Universal Robots URScript: FaiChun_9 Jan_7.script

def Machining1():
  # Default parameters:
  global speed_ms = 0.1
  global speed_rads = 0.75
  global accel_mss = 3
  global accel_radss = 1.2
  global blend_radius_m = 0.0002

  # Add subprograms here
  # Start of main program
  # Program generated by RoboDK v5.6.8 for UR10e on 10/01/2025 13:02:06
  # Using nominal kinematics.
  blend_radius_m = 0.0002
  speed_ms = 0.1
  # set_reference(p[0.355000, -0.055000, 0.001500, 0.000000, 0.000000, 0.000000])
  set_tcp(p[0.000000, 0.000000, 0.252000, 0.000000, 0.000000, 0.000000])
  # Show Tool
  movej([0.687885, -1.099321, -2.618738, -0.994329, 1.570796, 2.258681],accel_radss,speed_rads,0,blend_radius_m)
  movel([0.687885, -1.158787, -2.657718, -0.895884, 1.570796, 2.258681],accel_mss,speed_ms,0,blend_radius_m)
  #SetTool1
  #M_RunCode6
  #SetRPM60000
  speed_ms = 0.1
  #M_RunCode3
  movel([0.687885, -1.186172, -2.672546, -0.853671, 1.570796, 2.258681],accel_mss,speed_ms,0,blend_radius_m)
  speed_ms = 0.003
  movel([0.687885, -1.193386, -2.676190, -0.842813, 1.570796, 2.258681],accel_mss,speed_ms,0,blend_radius_m)
  speed_ms = 0.007
  movel([0.511185, -1.481281, -2.488242, -0.742866, 1.570796, 2.081982],accel_mss,speed_ms,0,blend_radius_m)
  movel([0.262250, -1.477063, -2.491849, -0.743477, 1.570796, 1.833046],accel_mss,speed_ms,0,blend_radius_m)
  movel([0.358500, -1.184451, -2.680352, -0.847585, 1.570796, 1.929297],accel_mss,speed_ms,0,blend_radius_m)
  movel([0.687885, -1.193386, -2.676190, -0.842813, 1.570796, 2.258681],accel_mss,speed_ms,0,blend_radius_m)
  speed_ms = 0.003
  movel([0.687885, -1.186172, -2.672546, -0.853671, 1.570796, 2.258681],accel_mss,speed_ms,0,blend_radius_m)
  speed_ms = 0.1
  movel([0.687885, -1.158787, -2.657718, -0.895884, 1.570796, 2.258681],accel_mss,speed_ms,0,blend_radius_m)
  #M_RunCode9
  movel([0.673659, -1.163346, -2.655655, -0.893388, 1.570796, 2.244455],accel_mss,speed_ms,0,blend_radius_m)
  #M_RunCode3
  movel([0.673659, -1.190701, -2.670423, -0.851265, 1.570796, 2.244455],accel_mss,speed_ms,0,blend_radius_m)
  speed_ms = 0.003
  movel([0.673659, -1.197905, -2.674052, -0.840433, 1.570796, 2.244455],accel_mss,speed_ms,0,blend_radius_m)
  speed_ms = 0.007
  movel([0.670159, -1.203367, -2.671437, -0.837585, 1.570796, 2.240955],accel_mss,speed_ms,0,blend_radius_m)
  movel([0.674542, -1.204354, -2.670961, -0.837074, 1.570796, 2.245338],accel_mss,speed_ms,0,blend_radius_m)
  movel([0.669404, -1.212334, -2.667074, -0.832981, 1.570796, 2.240200],accel_mss,speed_ms,0,blend_radius_m)
  movel([0.665043, -1.211367, -2.667549, -0.833473, 1.570796, 2.235840],accel_mss,speed_ms,0,blend_radius_m)
  movel([0.663268, -1.214147, -2.666181, -0.832061, 1.570796, 2.234065],accel_mss,speed_ms,0,blend_radius_m)
  movel([0.667621, -1.215107, -2.665706, -0.831575, 1.570796, 2.238418],accel_mss,speed_ms,0,blend_radius_m)
  movel([0.663402, -1.221682, -2.662429, -0.828278, 1.570796, 2.234198],accel_mss,speed_ms,0,blend_radius_m)
  movel([0.662590, -1.222948, -2.661792, -0.827649, 1.570796, 2.233387],accel_mss,speed_ms,0,blend_radius_m)
  movel([0.656171, -1.221563, -2.662488, -0.828337, 1.570796, 2.226968],accel_mss,speed_ms,0,blend_radius_m)
  movel([0.659538, -1.216260, -2.665135, -0.830994, 1.570796, 2.230334],accel_mss,speed_ms,0,blend_radius_m)
  movel([0.657269, -1.215780, -2.665373, -0.831236, 1.570796, 2.228065],accel_mss,speed_ms,0,blend_radius_m)
  movel([0.652180, -1.223829, -2.661348, -0.827212, 1.570796, 2.222977],accel_mss,speed_ms,0,blend_radius_m)
  movel([0.660845, -1.225674, -2.660415, -0.826300, 1.570796, 2.231641],accel_mss,speed_ms,0,blend_radius_m)
  movel([0.581204, -1.353206, -2.585789, -0.773394, 1.570796, 2.152000],accel_mss,speed_ms,0,blend_radius_m)
  movel([0.518903, -1.459211, -2.506807, -0.746371, 1.570796, 2.089699],accel_mss,speed_ms,0,blend_radius_m)
  movel([0.511689, -1.458211, -2.507631, -0.746547, 1.570796, 2.082486],accel_mss,speed_ms,0,blend_radius_m)
  movel([0.508628, -1.463700, -2.503092, -0.745597, 1.570796, 2.079424],accel_mss,speed_ms,0,blend_radius_m)
  movel([0.510492, -1.463952, -2.502883, -0.745554, 1.570796, 2.081288],accel_mss,speed_ms,0,blend_radius_m)
  movel([0.512509, -1.460346, -2.505871, -0.746172, 1.570796, 2.083305],accel_mss,speed_ms,0,blend_radius_m)
  movel([0.517829, -1.461092, -2.505254, -0.746043, 1.570796, 2.088625],accel_mss,speed_ms,0,blend_radius_m)
  movel([0.517338, -1.461959, -2.504537, -0.745893, 1.570796, 2.088135],accel_mss,speed_ms,0,blend_radius_m)
  movel([0.514822, -1.466415, -2.500830, -0.745144, 1.570796, 2.085618],accel_mss,speed_ms,0,blend_radius_m)
  movel([0.511249, -1.465915, -2.501248, -0.745226, 1.570796, 2.082045],accel_mss,speed_ms,0,blend_radius_m)
  movel([0.510209, -1.467774, -2.499694, -0.744921, 1.570796, 2.081005],accel_mss,speed_ms,0,blend_radius_m)
  movel([0.513778, -1.468272, -2.499276, -0.744840, 1.570796, 2.084574],accel_mss,speed_ms,0,blend_radius_m)
  movel([0.510816, -1.473540, -2.494840, -0.744009, 1.570796, 2.081613],accel_mss,speed_ms,0,blend_radius_m)
  movel([0.507266, -1.473049, -2.495255, -0.744085, 1.570796, 2.078063],accel_mss,speed_ms,0,blend_radius_m)
  movel([0.505298, -1.476588, -2.492253, -0.743548, 1.570796, 2.076095],accel_mss,speed_ms,0,blend_radius_m)
  movel([0.500042, -1.475891, -2.492846, -0.743652, 1.570796, 2.070838],accel_mss,speed_ms,0,blend_radius_m)
  movel([0.501993, -1.472345, -2.495850, -0.744194, 1.570796, 2.072789],accel_mss,speed_ms,0,blend_radius_m)
  movel([0.500139, -1.472105, -2.496053, -0.744231, 1.570796, 2.070935],accel_mss,speed_ms,0,blend_radius_m)
  movel([0.498194, -1.475653, -2.493048, -0.743688, 1.570796, 2.068990],accel_mss,speed_ms,0,blend_radius_m)
  movel([0.493769, -1.475101, -2.493517, -0.743771, 1.570796, 2.064565],accel_mss,speed_ms,0,blend_radius_m)
  movel([0.492911, -1.474994, -2.493608, -0.743787, 1.570796, 2.063707],accel_mss,speed_ms,0,blend_radius_m)
  movel([0.495770, -1.469725, -2.498057, -0.744607, 1.570796, 2.066567],accel_mss,speed_ms,0,blend_radius_m)
  movel([0.499358, -1.470173, -2.497681, -0.744536, 1.570796, 2.070154],accel_mss,speed_ms,0,blend_radius_m)
  movel([0.500375, -1.468318, -2.499238, -0.744833, 1.570796, 2.071171],accel_mss,speed_ms,0,blend_radius_m)
  movel([0.494912, -1.467639, -2.499806, -0.744943, 1.570796, 2.065708],accel_mss,speed_ms,0,blend_radius_m)
  movel([0.491053, -1.474772, -2.493796, -0.743821, 1.570796, 2.061849],accel_mss,speed_ms,0,blend_radius_m)
  movel([0.490192, -1.474669, -2.493883, -0.743837, 1.570796, 2.060989],accel_mss,speed_ms,0,blend_radius_m)
  movel([0.391239, -1.468060, -2.499454, -0.744875, 1.570796, 1.962036],accel_mss,speed_ms,0,blend_radius_m)
  movel([0.286918, -1.471352, -2.496688, -0.744349, 1.570796, 1.857714],accel_mss,speed_ms,0,blend_radius_m)
  movel([0.289237, -1.464153, -2.502716, -0.745520, 1.570796, 1.860034],accel_mss,speed_ms,0,blend_radius_m)
  movel([0.283249, -1.464641, -2.502309, -0.745438, 1.570796, 1.854046],accel_mss,speed_ms,0,blend_radius_m)
  movel([0.282655, -1.466514, -2.500748, -0.745128, 1.570796, 1.853451],accel_mss,speed_ms,0,blend_radius_m)
  movel([0.286590, -1.466190, -2.501018, -0.745181, 1.570796, 1.857386],accel_mss,speed_ms,0,blend_radius_m)
  movel([0.284883, -1.471507, -2.496557, -0.744325, 1.570796, 1.855679],accel_mss,speed_ms,0,blend_radius_m)
  movel([0.283941, -1.471581, -2.496494, -0.744313, 1.570796, 1.854738],accel_mss,speed_ms,0,blend_radius_m)
  movel([0.279090, -1.471983, -2.496155, -0.744250, 1.570796, 1.849887],accel_mss,speed_ms,0,blend_radius_m)
  movel([0.280215, -1.468402, -2.499167, -0.744819, 1.570796, 1.851011],accel_mss,speed_ms,0,blend_radius_m)
  movel([0.278175, -1.468578, -2.499020, -0.744791, 1.570796, 1.848972],accel_mss,speed_ms,0,blend_radius_m)
  movel([0.277057, -1.472158, -2.496008, -0.744223, 1.570796, 1.847854],accel_mss,speed_ms,0,blend_radius_m)
  movel([0.271256, -1.472675, -2.495571, -0.744143, 1.570796, 1.842052],accel_mss,speed_ms,0,blend_radius_m)
  movel([0.272350, -1.469100, -2.498582, -0.744707, 1.570796, 1.843147],accel_mss,speed_ms,0,blend_radius_m)
  movel([0.268413, -1.469469, -2.498272, -0.744648, 1.570796, 1.839210],accel_mss,speed_ms,0,blend_radius_m)
  movel([0.270027, -1.464147, -2.502721, -0.745521, 1.570796, 1.840824],accel_mss,speed_ms,0,blend_radius_m)
  movel([0.273986, -1.463773, -2.503032, -0.745584, 1.570796, 1.844782],accel_mss,speed_ms,0,blend_radius_m)
  movel([0.274565, -1.461897, -2.504588, -0.745904, 1.570796, 1.845361],accel_mss,speed_ms,0,blend_radius_m)
  movel([0.270596, -1.462271, -2.504279, -0.745840, 1.570796, 1.841392],accel_mss,speed_ms,0,blend_radius_m)
  movel([0.271969, -1.457770, -2.507994, -0.746626, 1.570796, 1.842765],accel_mss,speed_ms,0,blend_radius_m)
  movel([0.272236, -1.456894, -2.508713, -0.746782, 1.570796, 1.843033],accel_mss,speed_ms,0,blend_radius_m)
  movel([0.278152, -1.456332, -2.509173, -0.746883, 1.570796, 1.848948],accel_mss,speed_ms,0,blend_radius_m)
  movel([0.277017, -1.459975, -2.506178, -0.746237, 1.570796, 1.847813],accel_mss,speed_ms,0,blend_radius_m)
  movel([0.279080, -1.459787, -2.506332, -0.746270, 1.570796, 1.849877],accel_mss,speed_ms,0,blend_radius_m)
  movel([0.280818, -1.454246, -2.510881, -0.747263, 1.570796, 1.851615],accel_mss,speed_ms,0,blend_radius_m)
  movel([0.272819, -1.454995, -2.510268, -0.747126, 1.570796, 1.843616],accel_mss,speed_ms,0,blend_radius_m)
  movel([0.307084, -1.347659, -2.589476, -0.775253, 1.570796, 1.877880],accel_mss,speed_ms,0,blend_radius_m)
  movel([0.351247, -1.219193, -2.663675, -0.829521, 1.570796, 1.922043],accel_mss,speed_ms,0,blend_radius_m)
  movel([0.351702, -1.217910, -2.664315, -0.830164, 1.570796, 1.922499],accel_mss,speed_ms,0,blend_radius_m)
  movel([0.362053, -1.216508, -2.665012, -0.830869, 1.570796, 1.932849],accel_mss,speed_ms,0,blend_radius_m)
  movel([0.365050, -1.208304, -2.669046, -0.835039, 1.570796, 1.935846],accel_mss,speed_ms,0,blend_radius_m)
  movel([0.362345, -1.208664, -2.668871, -0.834855, 1.570796, 1.933142],accel_mss,speed_ms,0,blend_radius_m)
  movel([0.360382, -1.214071, -2.666218, -0.832100, 1.570796, 1.931178],accel_mss,speed_ms,0,blend_radius_m)
  movel([0.352706, -1.215118, -2.665701, -0.831570, 1.570796, 1.923502],accel_mss,speed_ms,0,blend_radius_m)
  movel([0.353163, -1.213827, -2.666339, -0.832224, 1.570796, 1.923959],accel_mss,speed_ms,0,blend_radius_m)
  movel([0.355556, -1.207116, -2.669624, -0.835649, 1.570796, 1.926352],accel_mss,speed_ms,0,blend_radius_m)
  movel([0.360785, -1.206388, -2.669977, -0.836024, 1.570796, 1.931582],accel_mss,speed_ms,0,blend_radius_m)
  movel([0.361812, -1.203551, -2.671348, -0.837489, 1.570796, 1.932609],accel_mss,speed_ms,0,blend_radius_m)
  movel([0.356568, -1.204285, -2.670995, -0.837109, 1.570796, 1.927364],accel_mss,speed_ms,0,blend_radius_m)
  movel([0.359487, -1.196137, -2.674891, -0.841361, 1.570796, 1.930283],accel_mss,speed_ms,0,blend_radius_m)
  movel([0.364775, -1.195388, -2.675245, -0.841756, 1.570796, 1.935572],accel_mss,speed_ms,0,blend_radius_m)
  movel([0.366805, -1.189812, -2.677865, -0.844712, 1.570796, 1.937602],accel_mss,speed_ms,0,blend_radius_m)
  movel([0.374669, -1.188736, -2.678367, -0.845286, 1.570796, 1.945465],accel_mss,speed_ms,0,blend_radius_m)
  movel([0.372594, -1.194327, -2.675746, -0.842316, 1.570796, 1.943391],accel_mss,speed_ms,0,blend_radius_m)
  movel([0.375333, -1.193969, -2.675915, -0.842505, 1.570796, 1.946129],accel_mss,speed_ms,0,blend_radius_m)
  movel([0.377422, -1.188372, -2.678536, -0.845481, 1.570796, 1.948219],accel_mss,speed_ms,0,blend_radius_m)
  movel([0.385265, -1.187376, -2.678999, -0.846014, 1.570796, 1.956062],accel_mss,speed_ms,0,blend_radius_m)
  movel([0.382115, -1.195666, -2.675114, -0.841609, 1.570796, 1.952912],accel_mss,speed_ms,0,blend_radius_m)
  movel([0.376864, -1.196318, -2.674805, -0.841266, 1.570796, 1.947660],accel_mss,speed_ms,0,blend_radius_m)
  movel([0.375787, -1.199193, -2.673438, -0.839758, 1.570796, 1.946584],accel_mss,speed_ms,0,blend_radius_m)
  movel([0.383743, -1.198220, -2.673902, -0.840267, 1.570796, 1.954539],accel_mss,speed_ms,0,blend_radius_m)
  movel([0.388012, -1.187041, -2.679154, -0.846193, 1.570796, 1.958808],accel_mss,speed_ms,0,blend_radius_m)
  movel([0.527415, -1.180130, -2.682335, -0.849924, 1.570796, 2.098211],accel_mss,speed_ms,0,blend_radius_m)
  movel([0.655859, -1.194143, -2.675833, -0.842413, 1.570796, 2.226656],accel_mss,speed_ms,0,blend_radius_m)
  movel([0.649023, -1.205134, -2.670585, -0.836671, 1.570796, 2.219819],accel_mss,speed_ms,0,blend_radius_m)
  movel([0.655771, -1.206472, -2.669937, -0.835981, 1.570796, 2.226568],accel_mss,speed_ms,0,blend_radius_m)
  movel([0.657545, -1.203650, -2.671301, -0.837438, 1.570796, 2.228341],accel_mss,speed_ms,0,blend_radius_m)
  movel([0.653099, -1.202756, -2.671731, -0.837902, 1.570796, 2.223896],accel_mss,speed_ms,0,blend_radius_m)
  movel([0.658190, -1.194618, -2.675609, -0.842162, 1.570796, 2.228986],accel_mss,speed_ms,0,blend_radius_m)
  movel([0.659266, -1.194835, -2.675507, -0.842048, 1.570796, 2.230062],accel_mss,speed_ms,0,blend_radius_m)
  movel([0.664798, -1.195978, -2.674966, -0.841445, 1.570796, 2.235595],accel_mss,speed_ms,0,blend_radius_m)
  movel([0.661332, -1.201468, -2.672350, -0.838571, 1.570796, 2.232128],accel_mss,speed_ms,0,blend_radius_m)
  movel([0.663629, -1.201951, -2.672118, -0.838320, 1.570796, 2.234425],accel_mss,speed_ms,0,blend_radius_m)
  movel([0.667108, -1.196468, -2.674734, -0.841187, 1.570796, 2.237905],accel_mss,speed_ms,0,blend_radius_m)
  movel([0.673659, -1.197905, -2.674052, -0.840433, 1.570796, 2.244455],accel_mss,speed_ms,0,blend_radius_m)
  speed_ms = 0.003
  movel([0.673659, -1.190701, -2.670423, -0.851265, 1.570796, 2.244455],accel_mss,speed_ms,0,blend_radius_m)
  speed_ms = 0.1
  movel([0.673659, -1.163346, -2.655655, -0.893388, 1.570796, 2.244455],accel_mss,speed_ms,0,blend_radius_m)
  #M_RunCode9
  movel([0.405490, -1.188907, -2.643693, -0.879789, 1.570796, 1.976287],accel_mss,speed_ms,0,blend_radius_m)
  #M_RunCode3
  movel([0.405490, -1.216061, -2.658125, -0.838204, 1.570796, 1.976287],accel_mss,speed_ms,0,blend_radius_m)
  speed_ms = 0.003
  movel([0.405490, -1.223196, -2.661667, -0.827526, 1.570796, 1.976287],accel_mss,speed_ms,0,blend_radius_m)
  speed_ms = 0.007
  movel([0.404235, -1.225666, -2.660419, -0.826304, 1.570796, 1.975032],accel_mss,speed_ms,0,blend_radius_m)
  movel([0.402333, -1.228061, -2.659202, -0.825126, 1.570796, 1.973129],accel_mss,speed_ms,0,blend_radius_m)
  movel([0.399790, -1.230382, -2.658016, -0.823990, 1.570796, 1.970587],accel_mss,speed_ms,0,blend_radius_m)
  movel([0.397246, -1.232154, -2.657107, -0.823128, 1.570796, 1.968043],accel_mss,speed_ms,0,blend_radius_m)
  movel([0.394666, -1.233434, -2.656448, -0.822507, 1.570796, 1.965462],accel_mss,speed_ms,0,blend_radius_m)
  movel([0.392112, -1.234311, -2.655995, -0.822083, 1.570796, 1.962908],accel_mss,speed_ms,0,blend_radius_m)
  movel([0.389658, -1.234867, -2.655708, -0.821814, 1.570796, 1.960454],accel_mss,speed_ms,0,blend_radius_m)
  movel([0.383823, -1.235506, -2.655377, -0.821506, 1.570796, 1.954620],accel_mss,speed_ms,0,blend_radius_m)
  movel([0.378293, -1.236171, -2.655032, -0.821186, 1.570796, 1.949089],accel_mss,speed_ms,0,blend_radius_m)
  movel([0.376058, -1.236689, -2.654763, -0.820937, 1.570796, 1.946854],accel_mss,speed_ms,0,blend_radius_m)
  movel([0.373771, -1.237485, -2.654349, -0.820555, 1.570796, 1.944568],accel_mss,speed_ms,0,blend_radius_m)
  movel([0.371510, -1.238623, -2.653756, -0.820010, 1.570796, 1.942306],accel_mss,speed_ms,0,blend_radius_m)
  movel([0.369355, -1.240154, -2.652956, -0.819279, 1.570796, 1.940152],accel_mss,speed_ms,0,blend_radius_m)
  movel([0.369832, -1.240875, -2.652578, -0.818936, 1.570796, 1.940628],accel_mss,speed_ms,0,blend_radius_m)
  movel([0.371300, -1.242746, -2.651595, -0.818048, 1.570796, 1.942096],accel_mss,speed_ms,0,blend_radius_m)
  movel([0.372894, -1.244134, -2.650863, -0.817392, 1.570796, 1.943691],accel_mss,speed_ms,0,blend_radius_m)
  movel([0.374621, -1.245036, -2.650386, -0.816967, 1.570796, 1.945417],accel_mss,speed_ms,0,blend_radius_m)
  movel([0.376480, -1.245459, -2.650162, -0.816768, 1.570796, 1.947276],accel_mss,speed_ms,0,blend_radius_m)
  movel([0.378426, -1.245454, -2.650164, -0.816771, 1.570796, 1.949222],accel_mss,speed_ms,0,blend_radius_m)
  movel([0.380419, -1.245079, -2.650363, -0.816947, 1.570796, 1.951216],accel_mss,speed_ms,0,blend_radius_m)
  movel([0.382465, -1.244329, -2.650760, -0.817300, 1.570796, 1.953261],accel_mss,speed_ms,0,blend_radius_m)
  movel([0.384565, -1.243203, -2.651354, -0.817832, 1.570796, 1.955361],accel_mss,speed_ms,0,blend_radius_m)
  movel([0.374982, -1.250934, -2.647243, -0.814212, 1.570796, 1.945778],accel_mss,speed_ms,0,blend_radius_m)
  movel([0.362201, -1.231769, -2.657305, -0.823315, 1.570796, 1.932997],accel_mss,speed_ms,0,blend_radius_m)
  movel([0.363171, -1.230958, -2.657721, -0.823709, 1.570796, 1.933967],accel_mss,speed_ms,0,blend_radius_m)
  movel([0.365784, -1.229122, -2.658661, -0.824606, 1.570796, 1.936581],accel_mss,speed_ms,0,blend_radius_m)
  movel([0.368660, -1.227763, -2.659354, -0.825272, 1.570796, 1.939456],accel_mss,speed_ms,0,blend_radius_m)
  movel([0.371629, -1.226820, -2.659834, -0.825736, 1.570796, 1.942425],accel_mss,speed_ms,0,blend_radius_m)
  movel([0.374540, -1.226217, -2.660140, -0.826032, 1.570796, 1.945337],accel_mss,speed_ms,0,blend_radius_m)
  movel([0.382124, -1.225371, -2.660568, -0.826449, 1.570796, 1.952921],accel_mss,speed_ms,0,blend_radius_m)
  movel([0.389118, -1.224702, -2.660907, -0.826780, 1.570796, 1.959914],accel_mss,speed_ms,0,blend_radius_m)
  movel([0.391824, -1.224204, -2.661159, -0.827026, 1.570796, 1.962621],accel_mss,speed_ms,0,blend_radius_m)
  movel([0.394534, -1.223409, -2.661560, -0.827420, 1.570796, 1.965331],accel_mss,speed_ms,0,blend_radius_m)
  movel([0.397109, -1.222267, -2.662135, -0.827987, 1.570796, 1.967906],accel_mss,speed_ms,0,blend_radius_m)
  movel([0.399421, -1.220716, -2.662914, -0.828760, 1.570796, 1.970217],accel_mss,speed_ms,0,blend_radius_m)
  movel([0.401837, -1.218360, -2.664091, -0.829938, 1.570796, 1.972633],accel_mss,speed_ms,0,blend_radius_m)
  movel([0.402665, -1.217183, -2.664677, -0.830529, 1.570796, 1.973461],accel_mss,speed_ms,0,blend_radius_m)
  movel([0.403233, -1.216010, -2.665259, -0.831120, 1.570796, 1.974029],accel_mss,speed_ms,0,blend_radius_m)
  movel([0.403673, -1.213869, -2.666318, -0.832202, 1.570796, 1.974470],accel_mss,speed_ms,0,blend_radius_m)
  movel([0.403233, -1.212154, -2.667162, -0.833073, 1.570796, 1.974029],accel_mss,speed_ms,0,blend_radius_m)
  movel([0.402520, -1.211325, -2.667569, -0.833495, 1.570796, 1.973317],accel_mss,speed_ms,0,blend_radius_m)
  movel([0.401656, -1.210987, -2.667735, -0.833667, 1.570796, 1.972453],accel_mss,speed_ms,0,blend_radius_m)
  movel([0.400727, -1.211098, -2.667681, -0.833611, 1.570796, 1.971523],accel_mss,speed_ms,0,blend_radius_m)
  movel([0.399832, -1.211610, -2.667429, -0.833349, 1.570796, 1.970628],accel_mss,speed_ms,0,blend_radius_m)
  movel([0.398841, -1.212924, -2.666784, -0.832682, 1.570796, 1.969637],accel_mss,speed_ms,0,blend_radius_m)
  movel([0.397954, -1.214245, -2.666132, -0.832012, 1.570796, 1.968750],accel_mss,speed_ms,0,blend_radius_m)
  movel([0.396541, -1.215617, -2.665454, -0.831318, 1.570796, 1.967337],accel_mss,speed_ms,0,blend_radius_m)
  movel([0.394622, -1.216822, -2.664856, -0.830711, 1.570796, 1.965418],accel_mss,speed_ms,0,blend_radius_m)
  movel([0.392868, -1.217184, -2.664676, -0.830529, 1.570796, 1.963664],accel_mss,speed_ms,0,blend_radius_m)
  movel([0.391414, -1.216814, -2.664860, -0.830715, 1.570796, 1.962211],accel_mss,speed_ms,0,blend_radius_m)
  movel([0.390392, -1.215820, -2.665353, -0.831216, 1.570796, 1.961188],accel_mss,speed_ms,0,blend_radius_m)
  movel([0.389911, -1.214381, -2.666065, -0.831943, 1.570796, 1.960708],accel_mss,speed_ms,0,blend_radius_m)
  movel([0.390088, -1.212670, -2.666908, -0.832810, 1.570796, 1.960884],accel_mss,speed_ms,0,blend_radius_m)
  movel([0.390972, -1.210867, -2.667794, -0.833728, 1.570796, 1.961769],accel_mss,speed_ms,0,blend_radius_m)
  movel([0.392610, -1.209162, -2.668628, -0.834599, 1.570796, 1.963406],accel_mss,speed_ms,0,blend_radius_m)
  movel([0.394268, -1.208010, -2.669189, -0.835190, 1.570796, 1.965064],accel_mss,speed_ms,0,blend_radius_m)
  movel([0.395903, -1.207293, -2.669538, -0.835558, 1.570796, 1.966700],accel_mss,speed_ms,0,blend_radius_m)
  movel([0.397515, -1.207013, -2.669674, -0.835702, 1.570796, 1.968311],accel_mss,speed_ms,0,blend_radius_m)
  movel([0.399100, -1.207171, -2.669597, -0.835621, 1.570796, 1.969897],accel_mss,speed_ms,0,blend_radius_m)
  movel([0.400597, -1.207720, -2.669330, -0.835339, 1.570796, 1.971394],accel_mss,speed_ms,0,blend_radius_m)
  movel([0.401956, -1.208596, -2.668904, -0.834890, 1.570796, 1.972752],accel_mss,speed_ms,0,blend_radius_m)
  movel([0.404240, -1.211338, -2.667563, -0.833488, 1.570796, 1.975036],accel_mss,speed_ms,0,blend_radius_m)
  movel([0.405266, -1.213469, -2.666515, -0.832405, 1.570796, 1.976062],accel_mss,speed_ms,0,blend_radius_m)
  movel([0.405912, -1.215735, -2.665395, -0.831258, 1.570796, 1.976709],accel_mss,speed_ms,0,blend_radius_m)
  movel([0.406187, -1.218131, -2.664205, -0.830053, 1.570796, 1.976983],accel_mss,speed_ms,0,blend_radius_m)
  movel([0.406094, -1.220651, -2.662946, -0.828792, 1.570796, 1.976890],accel_mss,speed_ms,0,blend_radius_m)
  movel([0.405490, -1.223196, -2.661667, -0.827526, 1.570796, 1.976287],accel_mss,speed_ms,0,blend_radius_m)
  speed_ms = 0.003
  movel([0.405490, -1.216061, -2.658125, -0.838204, 1.570796, 1.976287],accel_mss,speed_ms,0,blend_radius_m)
  speed_ms = 0.1
  movel([0.405490, -1.188907, -2.643693, -0.879789, 1.570796, 1.976287],accel_mss,speed_ms,0,blend_radius_m)
  #M_RunCode9
  movel([0.411128, -1.202346, -2.637125, -0.872918, 1.570796, 1.981924],accel_mss,speed_ms,0,blend_radius_m)
  #M_RunCode3
  movel([0.411128, -1.229375, -2.651380, -0.831635, 1.570796, 1.981924],accel_mss,speed_ms,0,blend_radius_m)
  speed_ms = 0.003
  movel([0.411128, -1.236469, -2.654877, -0.821043, 1.570796, 1.981924],accel_mss,speed_ms,0,blend_radius_m)
  speed_ms = 0.007
  movel([0.413224, -1.235399, -2.655432, -0.821558, 1.570796, 1.984020],accel_mss,speed_ms,0,blend_radius_m)
  movel([0.414871, -1.234902, -2.655690, -0.821797, 1.570796, 1.985668],accel_mss,speed_ms,0,blend_radius_m)
  movel([0.416069, -1.234980, -2.655649, -0.821760, 1.570796, 1.986865],accel_mss,speed_ms,0,blend_radius_m)
  movel([0.416819, -1.235628, -2.655314, -0.821447, 1.570796, 1.987615],accel_mss,speed_ms,0,blend_radius_m)
  movel([0.417031, -1.236693, -2.654761, -0.820935, 1.570796, 1.987827],accel_mss,speed_ms,0,blend_radius_m)
  movel([0.416624, -1.238016, -2.654073, -0.820300, 1.570796, 1.987421],accel_mss,speed_ms,0,blend_radius_m)
  movel([0.415599, -1.239598, -2.653247, -0.819544, 1.570796, 1.986395],accel_mss,speed_ms,0,blend_radius_m)
  movel([0.413957, -1.241437, -2.652283, -0.818669, 1.570796, 1.984754],accel_mss,speed_ms,0,blend_radius_m)
  movel([0.408873, -1.246069, -2.649839, -0.816482, 1.570796, 1.979669],accel_mss,speed_ms,0,blend_radius_m)
  movel([0.401436, -1.252092, -2.646621, -0.813676, 1.570796, 1.972233],accel_mss,speed_ms,0,blend_radius_m)
  movel([0.393892, -1.257776, -2.643545, -0.811068, 1.570796, 1.964688],accel_mss,speed_ms,0,blend_radius_m)
  movel([0.388401, -1.261422, -2.641551, -0.809415, 1.570796, 1.959198],accel_mss,speed_ms,0,blend_radius_m)
  movel([0.386373, -1.262468, -2.640976, -0.808945, 1.570796, 1.957169],accel_mss,speed_ms,0,blend_radius_m)
  movel([0.384770, -1.262965, -2.640703, -0.808721, 1.570796, 1.955566],accel_mss,speed_ms,0,blend_radius_m)
  movel([0.383590, -1.262914, -2.640731, -0.808744, 1.570796, 1.954386],accel_mss,speed_ms,0,blend_radius_m)
  movel([0.382828, -1.262317, -2.641059, -0.809012, 1.570796, 1.953624],accel_mss,speed_ms,0,blend_radius_m)
  movel([0.382577, -1.261314, -2.641611, -0.809464, 1.570796, 1.953374],accel_mss,speed_ms,0,blend_radius_m)
  movel([0.382928, -1.260047, -2.642305, -0.810037, 1.570796, 1.953725],accel_mss,speed_ms,0,blend_radius_m)
  movel([0.383890, -1.258512, -2.643144, -0.810733, 1.570796, 1.954686],accel_mss,speed_ms,0,blend_radius_m)
  movel([0.385460, -1.256708, -2.644126, -0.811555, 1.570796, 1.956257],accel_mss,speed_ms,0,blend_radius_m)
  movel([0.390413, -1.252101, -2.646616, -0.813672, 1.570796, 1.961210],accel_mss,speed_ms,0,blend_radius_m)
  movel([0.397814, -1.246023, -2.649863, -0.816503, 1.570796, 1.968610],accel_mss,speed_ms,0,blend_radius_m)
  movel([0.405474, -1.240218, -2.652923, -0.819249, 1.570796, 1.976271],accel_mss,speed_ms,0,blend_radius_m)
  movel([0.411128, -1.236469, -2.654877, -0.821043, 1.570796, 1.981924],accel_mss,speed_ms,0,blend_radius_m)
  speed_ms = 0.003
  movel([0.411128, -1.229375, -2.651380, -0.831635, 1.570796, 1.981924],accel_mss,speed_ms,0,blend_radius_m)
  speed_ms = 0.1
  movel([0.411128, -1.202346, -2.637125, -0.872918, 1.570796, 1.981924],accel_mss,speed_ms,0,blend_radius_m)
  #M_RunCode9
  movel([0.414372, -1.197750, -2.639394, -0.875246, 1.570796, 1.985169],accel_mss,speed_ms,0,blend_radius_m)
  #M_RunCode3
  movel([0.414372, -1.224822, -2.653709, -0.833858, 1.570796, 1.985169],accel_mss,speed_ms,0,blend_radius_m)
  speed_ms = 0.003
  movel([0.414372, -1.231931, -2.657222, -0.823236, 1.570796, 1.985169],accel_mss,speed_ms,0,blend_radius_m)
  speed_ms = 0.007
  movel([0.415723, -1.232648, -2.656853, -0.822888, 1.570796, 1.986520],accel_mss,speed_ms,0,blend_radius_m)
  movel([0.416849, -1.233640, -2.656342, -0.822407, 1.570796, 1.987645],accel_mss,speed_ms,0,blend_radius_m)
  movel([0.417744, -1.234908, -2.655686, -0.821794, 1.570796, 1.988541],accel_mss,speed_ms,0,blend_radius_m)
  movel([0.418377, -1.236379, -2.654924, -0.821086, 1.570796, 1.989173],accel_mss,speed_ms,0,blend_radius_m)
  movel([0.418708, -1.237979, -2.654092, -0.820318, 1.570796, 1.989504],accel_mss,speed_ms,0,blend_radius_m)
  movel([0.418737, -1.239713, -2.653187, -0.819489, 1.570796, 1.989533],accel_mss,speed_ms,0,blend_radius_m)
  movel([0.418470, -1.241571, -2.652213, -0.818605, 1.570796, 1.989266],accel_mss,speed_ms,0,blend_radius_m)
  movel([0.417892, -1.243534, -2.651180, -0.817675, 1.570796, 1.988689],accel_mss,speed_ms,0,blend_radius_m)
  movel([0.416999, -1.245570, -2.650103, -0.816716, 1.570796, 1.987795],accel_mss,speed_ms,0,blend_radius_m)
  movel([0.415789, -1.247678, -2.648983, -0.815728, 1.570796, 1.986585],accel_mss,speed_ms,0,blend_radius_m)
  movel([0.414266, -1.249863, -2.647817, -0.814709, 1.570796, 1.985063],accel_mss,speed_ms,0,blend_radius_m)
  movel([0.412445, -1.252075, -2.646630, -0.813684, 1.570796, 1.983241],accel_mss,speed_ms,0,blend_radius_m)
  movel([0.410340, -1.254273, -2.645445, -0.812671, 1.570796, 1.981136],accel_mss,speed_ms,0,blend_radius_m)
  movel([0.407956, -1.256457, -2.644262, -0.811669, 1.570796, 1.978752],accel_mss,speed_ms,0,blend_radius_m)
  movel([0.405287, -1.258633, -2.643078, -0.810678, 1.570796, 1.976084],accel_mss,speed_ms,0,blend_radius_m)
  movel([0.402539, -1.260646, -2.641977, -0.809766, 1.570796, 1.973335],accel_mss,speed_ms,0,blend_radius_m)
  movel([0.399900, -1.262345, -2.641044, -0.809000, 1.570796, 1.970696],accel_mss,speed_ms,0,blend_radius_m)
  movel([0.397372, -1.263737, -2.640277, -0.808375, 1.570796, 1.968168],accel_mss,speed_ms,0,blend_radius_m)
  movel([0.394950, -1.264822, -2.639678, -0.807889, 1.570796, 1.965746],accel_mss,speed_ms,0,blend_radius_m)
  movel([0.392670, -1.265602, -2.639246, -0.807541, 1.570796, 1.963466],accel_mss,speed_ms,0,blend_radius_m)
  movel([0.390566, -1.266088, -2.638976, -0.807325, 1.570796, 1.961362],accel_mss,speed_ms,0,blend_radius_m)
  movel([0.388636, -1.266279, -2.638870, -0.807240, 1.570796, 1.959432],accel_mss,speed_ms,0,blend_radius_m)
  movel([0.386882, -1.266174, -2.638928, -0.807286, 1.570796, 1.957678],accel_mss,speed_ms,0,blend_radius_m)
  movel([0.385319, -1.265788, -2.639143, -0.807458, 1.570796, 1.956115],accel_mss,speed_ms,0,blend_radius_m)
  movel([0.383964, -1.265145, -2.639499, -0.807745, 1.570796, 1.954760],accel_mss,speed_ms,0,blend_radius_m)
  movel([0.382821, -1.264237, -2.640001, -0.808151, 1.570796, 1.953617],accel_mss,speed_ms,0,blend_radius_m)
  movel([0.381888, -1.263063, -2.640649, -0.808677, 1.570796, 1.952684],accel_mss,speed_ms,0,blend_radius_m)
  movel([0.381205, -1.261689, -2.641405, -0.809295, 1.570796, 1.952002],accel_mss,speed_ms,0,blend_radius_m)
  movel([0.380815, -1.260177, -2.642234, -0.809978, 1.570796, 1.951611],accel_mss,speed_ms,0,blend_radius_m)
  movel([0.380719, -1.258521, -2.643139, -0.810729, 1.570796, 1.951515],accel_mss,speed_ms,0,blend_radius_m)
  movel([0.380920, -1.256723, -2.644118, -0.811548, 1.570796, 1.951717],accel_mss,speed_ms,0,blend_radius_m)
  movel([0.381427, -1.254806, -2.645157, -0.812426, 1.570796, 1.952224],accel_mss,speed_ms,0,blend_radius_m)
  movel([0.382253, -1.252799, -2.646241, -0.813349, 1.570796, 1.953050],accel_mss,speed_ms,0,blend_radius_m)
  movel([0.383399, -1.250697, -2.647370, -0.814322, 1.570796, 1.954196],accel_mss,speed_ms,0,blend_radius_m)
  movel([0.384868, -1.248499, -2.648545, -0.815344, 1.570796, 1.955664],accel_mss,speed_ms,0,blend_radius_m)
  movel([0.386648, -1.246250, -2.649742, -0.816397, 1.570796, 1.957444],accel_mss,speed_ms,0,blend_radius_m)
  movel([0.388736, -1.243991, -2.650938, -0.817460, 1.570796, 1.959532],accel_mss,speed_ms,0,blend_radius_m)
  movel([0.391132, -1.241721, -2.652134, -0.818534, 1.570796, 1.961928],accel_mss,speed_ms,0,blend_radius_m)
  movel([0.393832, -1.239446, -2.653326, -0.819617, 1.570796, 1.964629],accel_mss,speed_ms,0,blend_radius_m)
  movel([0.396644, -1.237322, -2.654434, -0.820633, 1.570796, 1.967441],accel_mss,speed_ms,0,blend_radius_m)
  movel([0.399357, -1.235518, -2.655371, -0.821500, 1.570796, 1.970154],accel_mss,speed_ms,0,blend_radius_m)
  movel([0.401972, -1.234038, -2.656136, -0.822215, 1.570796, 1.972769],accel_mss,speed_ms,0,blend_radius_m)
  movel([0.404484, -1.232879, -2.656734, -0.822776, 1.570796, 1.975280],accel_mss,speed_ms,0,blend_radius_m)
  movel([0.406847, -1.232048, -2.657162, -0.823179, 1.570796, 1.977643],accel_mss,speed_ms,0,blend_radius_m)
  movel([0.409023, -1.231537, -2.657424, -0.823428, 1.570796, 1.979819],accel_mss,speed_ms,0,blend_radius_m)
  movel([0.411005, -1.231352, -2.657519, -0.823518, 1.570796, 1.981802],accel_mss,speed_ms,0,blend_radius_m)
  movel([0.412793, -1.231491, -2.657448, -0.823450, 1.570796, 1.983589],accel_mss,speed_ms,0,blend_radius_m)
  movel([0.414372, -1.231931, -2.657222, -0.823236, 1.570796, 1.985169],accel_mss,speed_ms,0,blend_radius_m)
  speed_ms = 0.003
  movel([0.414372, -1.224822, -2.653709, -0.833858, 1.570796, 1.985169],accel_mss,speed_ms,0,blend_radius_m)
  speed_ms = 0.1
  movel([0.414372, -1.197750, -2.639394, -0.875246, 1.570796, 1.985169],accel_mss,speed_ms,0,blend_radius_m)
  #M_RunCode9
  movel([0.472103, -1.396064, -2.518448, -0.797877, 1.570796, 2.042899],accel_mss,speed_ms,0,blend_radius_m)
  #M_RunCode3
  movel([0.472103, -1.420124, -2.530197, -0.762068, 1.570796, 2.042899],accel_mss,speed_ms,0,blend_radius_m)
  speed_ms = 0.003
  movel([0.472103, -1.426356, -2.533062, -0.752970, 1.570796, 2.042899],accel_mss,speed_ms,0,blend_radius_m)
  speed_ms = 0.007
  movel([0.474230, -1.425319, -2.533865, -0.753205, 1.570796, 2.045026],accel_mss,speed_ms,0,blend_radius_m)
  movel([0.476498, -1.424700, -2.534343, -0.753346, 1.570796, 2.047294],accel_mss,speed_ms,0,blend_radius_m)
  movel([0.478796, -1.424421, -2.534558, -0.753410, 1.570796, 2.049593],accel_mss,speed_ms,0,blend_radius_m)
  movel([0.481016, -1.424399, -2.534575, -0.753415, 1.570796, 2.051812],accel_mss,speed_ms,0,blend_radius_m)
  movel([0.486722, -1.424913, -2.534179, -0.753298, 1.570796, 2.057518],accel_mss,speed_ms,0,blend_radius_m)
  movel([0.491970, -1.425464, -2.533753, -0.753172, 1.570796, 2.062767],accel_mss,speed_ms,0,blend_radius_m)
  movel([0.494023, -1.425488, -2.533734, -0.753167, 1.570796, 2.064819],accel_mss,speed_ms,0,blend_radius_m)
  movel([0.496103, -1.425282, -2.533893, -0.753214, 1.570796, 2.066899],accel_mss,speed_ms,0,blend_radius_m)
  movel([0.498116, -1.424785, -2.534277, -0.753327, 1.570796, 2.068912],accel_mss,speed_ms,0,blend_radius_m)
  movel([0.499969, -1.423929, -2.534937, -0.753523, 1.570796, 2.070765],accel_mss,speed_ms,0,blend_radius_m)
  movel([0.501973, -1.422467, -2.536063, -0.753860, 1.570796, 2.072769],accel_mss,speed_ms,0,blend_radius_m)
  movel([0.502690, -1.421679, -2.536667, -0.754042, 1.570796, 2.073486],accel_mss,speed_ms,0,blend_radius_m)
  movel([0.503217, -1.420854, -2.537300, -0.754235, 1.570796, 2.074014],accel_mss,speed_ms,0,blend_radius_m)
  movel([0.503737, -1.419264, -2.538516, -0.754609, 1.570796, 2.074534],accel_mss,speed_ms,0,blend_radius_m)
  movel([0.503565, -1.417868, -2.539581, -0.754940, 1.570796, 2.074361],accel_mss,speed_ms,0,blend_radius_m)
  movel([0.503117, -1.417117, -2.540153, -0.755120, 1.570796, 2.073913],accel_mss,speed_ms,0,blend_radius_m)
  movel([0.502508, -1.416723, -2.540452, -0.755214, 1.570796, 2.073304],accel_mss,speed_ms,0,blend_radius_m)
  movel([0.501814, -1.416665, -2.540496, -0.755228, 1.570796, 2.072610],accel_mss,speed_ms,0,blend_radius_m)
  movel([0.501105, -1.416925, -2.540299, -0.755166, 1.570796, 2.071901],accel_mss,speed_ms,0,blend_radius_m)
  movel([0.500253, -1.417791, -2.539640, -0.754959, 1.570796, 2.071049],accel_mss,speed_ms,0,blend_radius_m)
  movel([0.499479, -1.418679, -2.538962, -0.754747, 1.570796, 2.070275],accel_mss,speed_ms,0,blend_radius_m)
  movel([0.498307, -1.419527, -2.538315, -0.754547, 1.570796, 2.069103],accel_mss,speed_ms,0,blend_radius_m)
  movel([0.496779, -1.420169, -2.537825, -0.754396, 1.570796, 2.067575],accel_mss,speed_ms,0,blend_radius_m)
  movel([0.495450, -1.420178, -2.537817, -0.754393, 1.570796, 2.066246],accel_mss,speed_ms,0,blend_radius_m)
  movel([0.494407, -1.419666, -2.538209, -0.754514, 1.570796, 2.065204],accel_mss,speed_ms,0,blend_radius_m)
  movel([0.493744, -1.418737, -2.538918, -0.754733, 1.570796, 2.064540],accel_mss,speed_ms,0,blend_radius_m)
  movel([0.493526, -1.417542, -2.539829, -0.755018, 1.570796, 2.064322],accel_mss,speed_ms,0,blend_radius_m)
  movel([0.493817, -1.416240, -2.540819, -0.755330, 1.570796, 2.064613],accel_mss,speed_ms,0,blend_radius_m)
  movel([0.494639, -1.414976, -2.541777, -0.755636, 1.570796, 2.065435],accel_mss,speed_ms,0,blend_radius_m)
  movel([0.496006, -1.413907, -2.542586, -0.755896, 1.570796, 2.066803],accel_mss,speed_ms,0,blend_radius_m)
  movel([0.497336, -1.413272, -2.543066, -0.756051, 1.570796, 2.068132],accel_mss,speed_ms,0,blend_radius_m)
  movel([0.498607, -1.412968, -2.543295, -0.756126, 1.570796, 2.069403],accel_mss,speed_ms,0,blend_radius_m)
  movel([0.499820, -1.413002, -2.543270, -0.756118, 1.570796, 2.070616],accel_mss,speed_ms,0,blend_radius_m)
  movel([0.500972, -1.413373, -2.542990, -0.756027, 1.570796, 2.071769],accel_mss,speed_ms,0,blend_radius_m)
  movel([0.502028, -1.414027, -2.542495, -0.755866, 1.570796, 2.072825],accel_mss,speed_ms,0,blend_radius_m)
  movel([0.502947, -1.414917, -2.541822, -0.755650, 1.570796, 2.073743],accel_mss,speed_ms,0,blend_radius_m)
  movel([0.504384, -1.417391, -2.539944, -0.755054, 1.570796, 2.075180],accel_mss,speed_ms,0,blend_radius_m)
  movel([0.504947, -1.419197, -2.538567, -0.754625, 1.570796, 2.075743],accel_mss,speed_ms,0,blend_radius_m)
  movel([0.505221, -1.421051, -2.537149, -0.754189, 1.570796, 2.076017],accel_mss,speed_ms,0,blend_radius_m)
  movel([0.505212, -1.422947, -2.535694, -0.753749, 1.570796, 2.076008],accel_mss,speed_ms,0,blend_radius_m)
  movel([0.504914, -1.424889, -2.534197, -0.753303, 1.570796, 2.075711],accel_mss,speed_ms,0,blend_radius_m)
  movel([0.504239, -1.426773, -2.532739, -0.752876, 1.570796, 2.075036],accel_mss,speed_ms,0,blend_radius_m)
  movel([0.503088, -1.428504, -2.531396, -0.752489, 1.570796, 2.073884],accel_mss,speed_ms,0,blend_radius_m)
  movel([0.501463, -1.430083, -2.530167, -0.752140, 1.570796, 2.072259],accel_mss,speed_ms,0,blend_radius_m)
  movel([0.499365, -1.431510, -2.529052, -0.751827, 1.570796, 2.070162],accel_mss,speed_ms,0,blend_radius_m)
  movel([0.497315, -1.432509, -2.528270, -0.751610, 1.570796, 2.068112],accel_mss,speed_ms,0,blend_radius_m)
  movel([0.495279, -1.433123, -2.527788, -0.751478, 1.570796, 2.066075],accel_mss,speed_ms,0,blend_radius_m)
  movel([0.493299, -1.433425, -2.527551, -0.751412, 1.570796, 2.064095],accel_mss,speed_ms,0,blend_radius_m)
  movel([0.491422, -1.433491, -2.527499, -0.751398, 1.570796, 2.062218],accel_mss,speed_ms,0,blend_radius_m)
  movel([0.487019, -1.433111, -2.527798, -0.751480, 1.570796, 2.057815],accel_mss,speed_ms,0,blend_radius_m)
  movel([0.482843, -1.432791, -2.528049, -0.751549, 1.570796, 2.053639],accel_mss,speed_ms,0,blend_radius_m)
  movel([0.481129, -1.432857, -2.527997, -0.751535, 1.570796, 2.051925],accel_mss,speed_ms,0,blend_radius_m)
  movel([0.479349, -1.433136, -2.527778, -0.751475, 1.570796, 2.050145],accel_mss,speed_ms,0,blend_radius_m)
  movel([0.477553, -1.433686, -2.527347, -0.751356, 1.570796, 2.048350],accel_mss,speed_ms,0,blend_radius_m)
  movel([0.475798, -1.434563, -2.526657, -0.751169, 1.570796, 2.046594],accel_mss,speed_ms,0,blend_radius_m)
  movel([0.476083, -1.435203, -2.526154, -0.751033, 1.570796, 2.046880],accel_mss,speed_ms,0,blend_radius_m)
  movel([0.476995, -1.436904, -2.524811, -0.750673, 1.570796, 2.047791],accel_mss,speed_ms,0,blend_radius_m)
  movel([0.478051, -1.438239, -2.523755, -0.750395, 1.570796, 2.048847],accel_mss,speed_ms,0,blend_radius_m)
  movel([0.479252, -1.439214, -2.522982, -0.750193, 1.570796, 2.050048],accel_mss,speed_ms,0,blend_radius_m)
  movel([0.480597, -1.439828, -2.522495, -0.750066, 1.570796, 2.051393],accel_mss,speed_ms,0,blend_radius_m)
  movel([0.482052, -1.440117, -2.522265, -0.750007, 1.570796, 2.052848],accel_mss,speed_ms,0,blend_radius_m)
  movel([0.483576, -1.440121, -2.522262, -0.750006, 1.570796, 2.054373],accel_mss,speed_ms,0,blend_radius_m)
  movel([0.485174, -1.439838, -2.522487, -0.750064, 1.570796, 2.055971],accel_mss,speed_ms,0,blend_radius_m)
  movel([0.486848, -1.439266, -2.522941, -0.750182, 1.570796, 2.057644],accel_mss,speed_ms,0,blend_radius_m)
  movel([0.478951, -1.443924, -2.519227, -0.749238, 1.570796, 2.049747],accel_mss,speed_ms,0,blend_radius_m)
  movel([0.471303, -1.426844, -2.532684, -0.752861, 1.570796, 2.042099],accel_mss,speed_ms,0,blend_radius_m)
  movel([0.472103, -1.426356, -2.533062, -0.752970, 1.570796, 2.042899],accel_mss,speed_ms,0,blend_radius_m)
  speed_ms = 0.003
  movel([0.472103, -1.420124, -2.530197, -0.762068, 1.570796, 2.042899],accel_mss,speed_ms,0,blend_radius_m)
  speed_ms = 0.1
  movel([0.472103, -1.396064, -2.518448, -0.797877, 1.570796, 2.042899],accel_mss,speed_ms,0,blend_radius_m)
  #M_RunCode9
  movel([0.484799, -1.413284, -2.505502, -0.793604, 1.570796, 2.055595],accel_mss,speed_ms,0,blend_radius_m)
  #M_RunCode3
  movel([0.484799, -1.437005, -2.517040, -0.758344, 1.570796, 2.055595],accel_mss,speed_ms,0,blend_radius_m)
  speed_ms = 0.003
  movel([0.484799, -1.443143, -2.519852, -0.749394, 1.570796, 2.055595],accel_mss,speed_ms,0,blend_radius_m)
  speed_ms = 0.007
  movel([0.486288, -1.442519, -2.520351, -0.749519, 1.570796, 2.057084],accel_mss,speed_ms,0,blend_radius_m)
  movel([0.487606, -1.442497, -2.520368, -0.749523, 1.570796, 2.058403],accel_mss,speed_ms,0,blend_radius_m)
  movel([0.488644, -1.442984, -2.519979, -0.749426, 1.570796, 2.059440],accel_mss,speed_ms,0,blend_radius_m)
  movel([0.489301, -1.443881, -2.519261, -0.749246, 1.570796, 2.060098],accel_mss,speed_ms,0,blend_radius_m)
  movel([0.489515, -1.445038, -2.518334, -0.749017, 1.570796, 2.060311],accel_mss,speed_ms,0,blend_radius_m)
  movel([0.489218, -1.446300, -2.517321, -0.748769, 1.570796, 2.060014],accel_mss,speed_ms,0,blend_radius_m)
  movel([0.488417, -1.447511, -2.516345, -0.748533, 1.570796, 2.059213],accel_mss,speed_ms,0,blend_radius_m)
  movel([0.487104, -1.448523, -2.515528, -0.748338, 1.570796, 2.057900],accel_mss,speed_ms,0,blend_radius_m)
  movel([0.485874, -1.449086, -2.515073, -0.748230, 1.570796, 2.056671],accel_mss,speed_ms,0,blend_radius_m)
  movel([0.484850, -1.449267, -2.514927, -0.748195, 1.570796, 2.055647],accel_mss,speed_ms,0,blend_radius_m)
  movel([0.483799, -1.449529, -2.514715, -0.748145, 1.570796, 2.054595],accel_mss,speed_ms,0,blend_radius_m)
  movel([0.483225, -1.450019, -2.514318, -0.748052, 1.570796, 2.054021],accel_mss,speed_ms,0,blend_radius_m)
  movel([0.482865, -1.450694, -2.513771, -0.747924, 1.570796, 2.053661],accel_mss,speed_ms,0,blend_radius_m)
  movel([0.482750, -1.451433, -2.513171, -0.747785, 1.570796, 2.053546],accel_mss,speed_ms,0,blend_radius_m)
  movel([0.482905, -1.452122, -2.512611, -0.747656, 1.570796, 2.053701],accel_mss,speed_ms,0,blend_radius_m)
  movel([0.483377, -1.452876, -2.511998, -0.747516, 1.570796, 2.054173],accel_mss,speed_ms,0,blend_radius_m)
  movel([0.484052, -1.453420, -2.511554, -0.747415, 1.570796, 2.054849],accel_mss,speed_ms,0,blend_radius_m)
  movel([0.484931, -1.453757, -2.511280, -0.747353, 1.570796, 2.055727],accel_mss,speed_ms,0,blend_radius_m)
  movel([0.486011, -1.453886, -2.511174, -0.747329, 1.570796, 2.056807],accel_mss,speed_ms,0,blend_radius_m)
  movel([0.487228, -1.453801, -2.511243, -0.747344, 1.570796, 2.058025],accel_mss,speed_ms,0,blend_radius_m)
  movel([0.488523, -1.453496, -2.511492, -0.747401, 1.570796, 2.059319],accel_mss,speed_ms,0,blend_radius_m)
  movel([0.489895, -1.452968, -2.511923, -0.747498, 1.570796, 2.060691],accel_mss,speed_ms,0,blend_radius_m)
  movel([0.491344, -1.452220, -2.512532, -0.747637, 1.570796, 2.062140],accel_mss,speed_ms,0,blend_radius_m)
  movel([0.493609, -1.450595, -2.513851, -0.747943, 1.570796, 2.064406],accel_mss,speed_ms,0,blend_radius_m)
  movel([0.495423, -1.448595, -2.515470, -0.748324, 1.570796, 2.066219],accel_mss,speed_ms,0,blend_radius_m)
  movel([0.496139, -1.447461, -2.516386, -0.748543, 1.570796, 2.066936],accel_mss,speed_ms,0,blend_radius_m)
  movel([0.496696, -1.446248, -2.517362, -0.748779, 1.570796, 2.067492],accel_mss,speed_ms,0,blend_radius_m)
  movel([0.497331, -1.443593, -2.519493, -0.749304, 1.570796, 2.068127],accel_mss,speed_ms,0,blend_radius_m)
  movel([0.497249, -1.440695, -2.521806, -0.749889, 1.570796, 2.068045],accel_mss,speed_ms,0,blend_radius_m)
  movel([0.496363, -1.437639, -2.524230, -0.750520, 1.570796, 2.067160],accel_mss,speed_ms,0,blend_radius_m)
  movel([0.508638, -1.430570, -2.529786, -0.752033, 1.570796, 2.079434],accel_mss,speed_ms,0,blend_radius_m)
  movel([0.513717, -1.443743, -2.519372, -0.749274, 1.570796, 2.084514],accel_mss,speed_ms,0,blend_radius_m)
  movel([0.505802, -1.448207, -2.515784, -0.748398, 1.570796, 2.076598],accel_mss,speed_ms,0,blend_radius_m)
  movel([0.507494, -1.446644, -2.517044, -0.748701, 1.570796, 2.078291],accel_mss,speed_ms,0,blend_radius_m)
  movel([0.508859, -1.444763, -2.518555, -0.749071, 1.570796, 2.079655],accel_mss,speed_ms,0,blend_radius_m)
  movel([0.509823, -1.442651, -2.520246, -0.749493, 1.570796, 2.080619],accel_mss,speed_ms,0,blend_radius_m)
  movel([0.510316, -1.440405, -2.522036, -0.749948, 1.570796, 2.081112],accel_mss,speed_ms,0,blend_radius_m)
  movel([0.510294, -1.438111, -2.523857, -0.750421, 1.570796, 2.081091],accel_mss,speed_ms,0,blend_radius_m)
  movel([0.509713, -1.435861, -2.525635, -0.750893, 1.570796, 2.080509],accel_mss,speed_ms,0,blend_radius_m)
  movel([0.500686, -1.441018, -2.521548, -0.749823, 1.570796, 2.071483],accel_mss,speed_ms,0,blend_radius_m)
  movel([0.501475, -1.443733, -2.519381, -0.749276, 1.570796, 2.072271],accel_mss,speed_ms,0,blend_radius_m)
  movel([0.501719, -1.446615, -2.517067, -0.748707, 1.570796, 2.072516],accel_mss,speed_ms,0,blend_radius_m)
  movel([0.501334, -1.449510, -2.514730, -0.748149, 1.570796, 2.072130],accel_mss,speed_ms,0,blend_radius_m)
  movel([0.500867, -1.450907, -2.513598, -0.747884, 1.570796, 2.071664],accel_mss,speed_ms,0,blend_radius_m)
  movel([0.500223, -1.452273, -2.512488, -0.747628, 1.570796, 2.071019],accel_mss,speed_ms,0,blend_radius_m)
  movel([0.499382, -1.453563, -2.511437, -0.747388, 1.570796, 2.070178],accel_mss,speed_ms,0,blend_radius_m)
  movel([0.498328, -1.454744, -2.510474, -0.747172, 1.570796, 2.069124],accel_mss,speed_ms,0,blend_radius_m)
  movel([0.497065, -1.455812, -2.509600, -0.746977, 1.570796, 2.067861],accel_mss,speed_ms,0,blend_radius_m)
  movel([0.495590, -1.456770, -2.508814, -0.746804, 1.570796, 2.066387],accel_mss,speed_ms,0,blend_radius_m)
  movel([0.494040, -1.457549, -2.508175, -0.746665, 1.570796, 2.064836],accel_mss,speed_ms,0,blend_radius_m)
  movel([0.492549, -1.458080, -2.507738, -0.746570, 1.570796, 2.063345],accel_mss,speed_ms,0,blend_radius_m)
  movel([0.491119, -1.458365, -2.507504, -0.746520, 1.570796, 2.061916],accel_mss,speed_ms,0,blend_radius_m)
  movel([0.489745, -1.458405, -2.507471, -0.746513, 1.570796, 2.060541],accel_mss,speed_ms,0,blend_radius_m)
  movel([0.487252, -1.457896, -2.507890, -0.746603, 1.570796, 2.058048],accel_mss,speed_ms,0,blend_radius_m)
  movel([0.485155, -1.456703, -2.508869, -0.746817, 1.570796, 2.055951],accel_mss,speed_ms,0,blend_radius_m)
  movel([0.483485, -1.454991, -2.510271, -0.747126, 1.570796, 2.054281],accel_mss,speed_ms,0,blend_radius_m)
  movel([0.482277, -1.452928, -2.511955, -0.747506, 1.570796, 2.053073],accel_mss,speed_ms,0,blend_radius_m)
  movel([0.481775, -1.451321, -2.513262, -0.747806, 1.570796, 2.052572],accel_mss,speed_ms,0,blend_radius_m)
  movel([0.481584, -1.449505, -2.514734, -0.748150, 1.570796, 2.052380],accel_mss,speed_ms,0,blend_radius_m)
  movel([0.481750, -1.447636, -2.516245, -0.748509, 1.570796, 2.052546],accel_mss,speed_ms,0,blend_radius_m)
  movel([0.482333, -1.445858, -2.517676, -0.748855, 1.570796, 2.053129],accel_mss,speed_ms,0,blend_radius_m)
  movel([0.483342, -1.444316, -2.518913, -0.749160, 1.570796, 2.054139],accel_mss,speed_ms,0,blend_radius_m)
  movel([0.484799, -1.443143, -2.519852, -0.749394, 1.570796, 2.055595],accel_mss,speed_ms,0,blend_radius_m)
  speed_ms = 0.003
  movel([0.484799, -1.437005, -2.517040, -0.758344, 1.570796, 2.055595],accel_mss,speed_ms,0,blend_radius_m)
  speed_ms = 0.1
  movel([0.484799, -1.413284, -2.505502, -0.793604, 1.570796, 2.055595],accel_mss,speed_ms,0,blend_radius_m)
  #M_RunCode9
  movel([0.488437, -1.342214, -2.556269, -0.813905, 1.570796, 2.059233],accel_mss,speed_ms,0,blend_radius_m)
  #M_RunCode3
  movel([0.488437, -1.367276, -2.568695, -0.776418, 1.570796, 2.059233],accel_mss,speed_ms,0,blend_radius_m)
  speed_ms = 0.003
  movel([0.488437, -1.373788, -2.571730, -0.766870, 1.570796, 2.059233],accel_mss,speed_ms,0,blend_radius_m)
  speed_ms = 0.007
  movel([0.485960, -1.374281, -2.571387, -0.766722, 1.570796, 2.056756],accel_mss,speed_ms,0,blend_radius_m)
  movel([0.483541, -1.374282, -2.571386, -0.766721, 1.570796, 2.054337],accel_mss,speed_ms,0,blend_radius_m)
  movel([0.481234, -1.373869, -2.571674, -0.766846, 1.570796, 2.052030],accel_mss,speed_ms,0,blend_radius_m)
  movel([0.479095, -1.373128, -2.572191, -0.767070, 1.570796, 2.049891],accel_mss,speed_ms,0,blend_radius_m)
  movel([0.477178, -1.372136, -2.572881, -0.767372, 1.570796, 2.047975],accel_mss,speed_ms,0,blend_radius_m)
  movel([0.478516, -1.369320, -2.574833, -0.768236, 1.570796, 2.049312],accel_mss,speed_ms,0,blend_radius_m)
  movel([0.480669, -1.366302, -2.576913, -0.769174, 1.570796, 2.051465],accel_mss,speed_ms,0,blend_radius_m)
  movel([0.483411, -1.363356, -2.578930, -0.770103, 1.570796, 2.054208],accel_mss,speed_ms,0,blend_radius_m)
  movel([0.486513, -1.360759, -2.580699, -0.770931, 1.570796, 2.057309],accel_mss,speed_ms,0,blend_radius_m)
  movel([0.489731, -1.358793, -2.582031, -0.771565, 1.570796, 2.060527],accel_mss,speed_ms,0,blend_radius_m)
  movel([0.491307, -1.358136, -2.582475, -0.771777, 1.570796, 2.062103],accel_mss,speed_ms,0,blend_radius_m)
  movel([0.492819, -1.357746, -2.582739, -0.771904, 1.570796, 2.063616],accel_mss,speed_ms,0,blend_radius_m)
  movel([0.494240, -1.357652, -2.582802, -0.771935, 1.570796, 2.065036],accel_mss,speed_ms,0,blend_radius_m)
  movel([0.495532, -1.357896, -2.582638, -0.771856, 1.570796, 2.066329],accel_mss,speed_ms,0,blend_radius_m)
  movel([0.496668, -1.358506, -2.582225, -0.771657, 1.570796, 2.067464],accel_mss,speed_ms,0,blend_radius_m)
  movel([0.497617, -1.359519, -2.581540, -0.771330, 1.570796, 2.068413],accel_mss,speed_ms,0,blend_radius_m)
  movel([0.498367, -1.361469, -2.580216, -0.770704, 1.570796, 2.069163],accel_mss,speed_ms,0,blend_radius_m)
  movel([0.498228, -1.363674, -2.578713, -0.770002, 1.570796, 2.069025],accel_mss,speed_ms,0,blend_radius_m)
  movel([0.497306, -1.366042, -2.577091, -0.769256, 1.570796, 2.068102],accel_mss,speed_ms,0,blend_radius_m)
  movel([0.495698, -1.368480, -2.575413, -0.768496, 1.570796, 2.066494],accel_mss,speed_ms,0,blend_radius_m)
  movel([0.493358, -1.370977, -2.573686, -0.767726, 1.570796, 2.064154],accel_mss,speed_ms,0,blend_radius_m)
  movel([0.490920, -1.372715, -2.572478, -0.767196, 1.570796, 2.061716],accel_mss,speed_ms,0,blend_radius_m)
  movel([0.488437, -1.373788, -2.571730, -0.766870, 1.570796, 2.059233],accel_mss,speed_ms,0,blend_radius_m)
  speed_ms = 0.003
  movel([0.488437, -1.367276, -2.568695, -0.776418, 1.570796, 2.059233],accel_mss,speed_ms,0,blend_radius_m)
  speed_ms = 0.1
  movel([0.488437, -1.342214, -2.556269, -0.813905, 1.570796, 2.059233],accel_mss,speed_ms,0,blend_radius_m)
  #M_RunCode9
  movel([0.559176, -1.266608, -2.602919, -0.842862, 1.570796, 2.129973],accel_mss,speed_ms,0,blend_radius_m)
  #M_RunCode3
  movel([0.559176, -1.292870, -2.616326, -0.803193, 1.570796, 2.129973],accel_mss,speed_ms,0,blend_radius_m)
  speed_ms = 0.003
  movel([0.559176, -1.299730, -2.619609, -0.793051, 1.570796, 2.129973],accel_mss,speed_ms,0,blend_radius_m)
  speed_ms = 0.007
  movel([0.558187, -1.298790, -2.620169, -0.793430, 1.570796, 2.128983],accel_mss,speed_ms,0,blend_radius_m)
  movel([0.557585, -1.297494, -2.620940, -0.793955, 1.570796, 2.128381],accel_mss,speed_ms,0,blend_radius_m)
  movel([0.557205, -1.296013, -2.621819, -0.794557, 1.570796, 2.128001],accel_mss,speed_ms,0,blend_radius_m)
  movel([0.557916, -1.295811, -2.621938, -0.794640, 1.570796, 2.128713],accel_mss,speed_ms,0,blend_radius_m)
  movel([0.558340, -1.296094, -2.621771, -0.794524, 1.570796, 2.129137],accel_mss,speed_ms,0,blend_radius_m)
  movel([0.558868, -1.296379, -2.621602, -0.794408, 1.570796, 2.129664],accel_mss,speed_ms,0,blend_radius_m)
  movel([0.559895, -1.296178, -2.621721, -0.794490, 1.570796, 2.130691],accel_mss,speed_ms,0,blend_radius_m)
  movel([0.561027, -1.295534, -2.622102, -0.794753, 1.570796, 2.131823],accel_mss,speed_ms,0,blend_radius_m)
  movel([0.562109, -1.294692, -2.622600, -0.795097, 1.570796, 2.132905],accel_mss,speed_ms,0,blend_radius_m)
  movel([0.563586, -1.293481, -2.623314, -0.795594, 1.570796, 2.134383],accel_mss,speed_ms,0,blend_radius_m)
  movel([0.563232, -1.291547, -2.624451, -0.796391, 1.570796, 2.134028],accel_mss,speed_ms,0,blend_radius_m)
  movel([0.562354, -1.290296, -2.625184, -0.796909, 1.570796, 2.133150],accel_mss,speed_ms,0,blend_radius_m)
  movel([0.561669, -1.290022, -2.625344, -0.797023, 1.570796, 2.132466],accel_mss,speed_ms,0,blend_radius_m)
  movel([0.560796, -1.290036, -2.625336, -0.797017, 1.570796, 2.131593],accel_mss,speed_ms,0,blend_radius_m)
  movel([0.559714, -1.290374, -2.625138, -0.796877, 1.570796, 2.130510],accel_mss,speed_ms,0,blend_radius_m)
  movel([0.558409, -1.291077, -2.624726, -0.796585, 1.570796, 2.129206],accel_mss,speed_ms,0,blend_radius_m)
  movel([0.558885, -1.289731, -2.625514, -0.797144, 1.570796, 2.129681],accel_mss,speed_ms,0,blend_radius_m)
  movel([0.559453, -1.288575, -2.626189, -0.797625, 1.570796, 2.130249],accel_mss,speed_ms,0,blend_radius_m)
  movel([0.559811, -1.288164, -2.626428, -0.797797, 1.570796, 2.130608],accel_mss,speed_ms,0,blend_radius_m)
  movel([0.560236, -1.287918, -2.626571, -0.797900, 1.570796, 2.131033],accel_mss,speed_ms,0,blend_radius_m)
  movel([0.561357, -1.288072, -2.626481, -0.797835, 1.570796, 2.132153],accel_mss,speed_ms,0,blend_radius_m)
  movel([0.563064, -1.289295, -2.625769, -0.797325, 1.570796, 2.133861],accel_mss,speed_ms,0,blend_radius_m)
  movel([0.564262, -1.291053, -2.624741, -0.796595, 1.570796, 2.135059],accel_mss,speed_ms,0,blend_radius_m)
  movel([0.564539, -1.292099, -2.624127, -0.796163, 1.570796, 2.135336],accel_mss,speed_ms,0,blend_radius_m)
  movel([0.564531, -1.293236, -2.623458, -0.795695, 1.570796, 2.135328],accel_mss,speed_ms,0,blend_radius_m)
  movel([0.564188, -1.294448, -2.622744, -0.795197, 1.570796, 2.134984],accel_mss,speed_ms,0,blend_radius_m)
  movel([0.563456, -1.295725, -2.621989, -0.794675, 1.570796, 2.134252],accel_mss,speed_ms,0,blend_radius_m)
  movel([0.562339, -1.295007, -2.622414, -0.794968, 1.570796, 2.133135],accel_mss,speed_ms,0,blend_radius_m)
  movel([0.560715, -1.300130, -2.619369, -0.792889, 1.570796, 2.131512],accel_mss,speed_ms,0,blend_radius_m)
  movel([0.559176, -1.299730, -2.619609, -0.793051, 1.570796, 2.129973],accel_mss,speed_ms,0,blend_radius_m)
  speed_ms = 0.003
  movel([0.559176, -1.292870, -2.616326, -0.803193, 1.570796, 2.129973],accel_mss,speed_ms,0,blend_radius_m)
  speed_ms = 0.1
  movel([0.559176, -1.266608, -2.602919, -0.842862, 1.570796, 2.129973],accel_mss,speed_ms,0,blend_radius_m)
  #M_RunCode9
  movel([0.541155, -1.231973, -2.621944, -0.858472, 1.570796, 2.111951],accel_mss,speed_ms,0,blend_radius_m)
  #M_RunCode3
  movel([0.541155, -1.258681, -2.635807, -0.817901, 1.570796, 2.111951],accel_mss,speed_ms,0,blend_radius_m)
  speed_ms = 0.003
  movel([0.541155, -1.265675, -2.639205, -0.807509, 1.570796, 2.111951],accel_mss,speed_ms,0,blend_radius_m)
  speed_ms = 0.007
  movel([0.538885, -1.267349, -2.638276, -0.806764, 1.570796, 2.109681],accel_mss,speed_ms,0,blend_radius_m)
  movel([0.536503, -1.268835, -2.637448, -0.806106, 1.570796, 2.107299],accel_mss,speed_ms,0,blend_radius_m)
  movel([0.534036, -1.270098, -2.636742, -0.805549, 1.570796, 2.104832],accel_mss,speed_ms,0,blend_radius_m)
  movel([0.531508, -1.271114, -2.636173, -0.805102, 1.570796, 2.102304],accel_mss,speed_ms,0,blend_radius_m)
  movel([0.528945, -1.271858, -2.635755, -0.804776, 1.570796, 2.099741],accel_mss,speed_ms,0,blend_radius_m)
  movel([0.527649, -1.271977, -2.635688, -0.804724, 1.570796, 2.098445],accel_mss,speed_ms,0,blend_radius_m)
  movel([0.526355, -1.271896, -2.635734, -0.804759, 1.570796, 2.097151],accel_mss,speed_ms,0,blend_radius_m)
  movel([0.525190, -1.271832, -2.635770, -0.804787, 1.570796, 2.095986],accel_mss,speed_ms,0,blend_radius_m)
  movel([0.524282, -1.271998, -2.635677, -0.804715, 1.570796, 2.095078],accel_mss,speed_ms,0,blend_radius_m)
  movel([0.522755, -1.273059, -2.635079, -0.804250, 1.570796, 2.093551],accel_mss,speed_ms,0,blend_radius_m)
  movel([0.520756, -1.274766, -2.634116, -0.803507, 1.570796, 2.091553],accel_mss,speed_ms,0,blend_radius_m)
  movel([0.518685, -1.276566, -2.633096, -0.802727, 1.570796, 2.089481],accel_mss,speed_ms,0,blend_radius_m)
  movel([0.516926, -1.277918, -2.632328, -0.802143, 1.570796, 2.087722],accel_mss,speed_ms,0,blend_radius_m)
  movel([0.513420, -1.279914, -2.631189, -0.801286, 1.570796, 2.084217],accel_mss,speed_ms,0,blend_radius_m)
  movel([0.510269, -1.281209, -2.630447, -0.800733, 1.570796, 2.081065],accel_mss,speed_ms,0,blend_radius_m)
  movel([0.507438, -1.281868, -2.630069, -0.800452, 1.570796, 2.078235],accel_mss,speed_ms,0,blend_radius_m)
  movel([0.504899, -1.281960, -2.630016, -0.800413, 1.570796, 2.075696],accel_mss,speed_ms,0,blend_radius_m)
  movel([0.502627, -1.281549, -2.630252, -0.800588, 1.570796, 2.073423],accel_mss,speed_ms,0,blend_radius_m)
  movel([0.500595, -1.280695, -2.630742, -0.800952, 1.570796, 2.071391],accel_mss,speed_ms,0,blend_radius_m)
  movel([0.498776, -1.279468, -2.631444, -0.801478, 1.570796, 2.069572],accel_mss,speed_ms,0,blend_radius_m)
  movel([0.497148, -1.277921, -2.632326, -0.802142, 1.570796, 2.067944],accel_mss,speed_ms,0,blend_radius_m)
  movel([0.494376, -1.274127, -2.634477, -0.803785, 1.570796, 2.065172],accel_mss,speed_ms,0,blend_radius_m)
  movel([0.492091, -1.269821, -2.636897, -0.805671, 1.570796, 2.062888],accel_mss,speed_ms,0,blend_radius_m)
  movel([0.488292, -1.261723, -2.641386, -0.809280, 1.570796, 2.059088],accel_mss,speed_ms,0,blend_radius_m)
  movel([0.486181, -1.258480, -2.643161, -0.810748, 1.570796, 2.056977],accel_mss,speed_ms,0,blend_radius_m)
  movel([0.483296, -1.255078, -2.645010, -0.812301, 1.570796, 2.054092],accel_mss,speed_ms,0,blend_radius_m)
  movel([0.479761, -1.251728, -2.646817, -0.813844, 1.570796, 2.050558],accel_mss,speed_ms,0,blend_radius_m)
  movel([0.475699, -1.248636, -2.648473, -0.815281, 1.570796, 2.046495],accel_mss,speed_ms,0,blend_radius_m)
  movel([0.471246, -1.246011, -2.649869, -0.816509, 1.570796, 2.042042],accel_mss,speed_ms,0,blend_radius_m)
  movel([0.466543, -1.244058, -2.650903, -0.817428, 1.570796, 2.037339],accel_mss,speed_ms,0,blend_radius_m)
  movel([0.461738, -1.242979, -2.651472, -0.817938, 1.570796, 2.032535],accel_mss,speed_ms,0,blend_radius_m)
  movel([0.459347, -1.242827, -2.651552, -0.818010, 1.570796, 2.030144],accel_mss,speed_ms,0,blend_radius_m)
  movel([0.456991, -1.242963, -2.651480, -0.817945, 1.570796, 2.027788],accel_mss,speed_ms,0,blend_radius_m)
  movel([0.454465, -1.243412, -2.651244, -0.817733, 1.570796, 2.025261],accel_mss,speed_ms,0,blend_radius_m)
  movel([0.451439, -1.244221, -2.650817, -0.817351, 1.570796, 2.022236],accel_mss,speed_ms,0,blend_radius_m)
  movel([0.448094, -1.245409, -2.650188, -0.816792, 1.570796, 2.018890],accel_mss,speed_ms,0,blend_radius_m)
  movel([0.444604, -1.246992, -2.649348, -0.816049, 1.570796, 2.015400],accel_mss,speed_ms,0,blend_radius_m)
  movel([0.441140, -1.248986, -2.648286, -0.815118, 1.570796, 2.011937],accel_mss,speed_ms,0,blend_radius_m)
  movel([0.437888, -1.251398, -2.646994, -0.813997, 1.570796, 2.008684],accel_mss,speed_ms,0,blend_radius_m)
  movel([0.435011, -1.254243, -2.645461, -0.812684, 1.570796, 2.005808],accel_mss,speed_ms,0,blend_radius_m)
  movel([0.433772, -1.255826, -2.644605, -0.811958, 1.570796, 2.004569],accel_mss,speed_ms,0,blend_radius_m)
  movel([0.432693, -1.257522, -2.643683, -0.811184, 1.570796, 2.003489],accel_mss,speed_ms,0,blend_radius_m)
  movel([0.431527, -1.260176, -2.642234, -0.809978, 1.570796, 2.002323],accel_mss,speed_ms,0,blend_radius_m)
  movel([0.431211, -1.262432, -2.640996, -0.808961, 1.570796, 2.002007],accel_mss,speed_ms,0,blend_radius_m)
  movel([0.431652, -1.264327, -2.639952, -0.808111, 1.570796, 2.002448],accel_mss,speed_ms,0,blend_radius_m)
  movel([0.432753, -1.265897, -2.639082, -0.807410, 1.570796, 2.003550],accel_mss,speed_ms,0,blend_radius_m)
  movel([0.434427, -1.267180, -2.638370, -0.806839, 1.570796, 2.005224],accel_mss,speed_ms,0,blend_radius_m)
  movel([0.436577, -1.268210, -2.637796, -0.806382, 1.570796, 2.007373],accel_mss,speed_ms,0,blend_radius_m)
  movel([0.439116, -1.269027, -2.637341, -0.806021, 1.570796, 2.009913],accel_mss,speed_ms,0,blend_radius_m)
  movel([0.441951, -1.269659, -2.636988, -0.805742, 1.570796, 2.012747],accel_mss,speed_ms,0,blend_radius_m)
  movel([0.448166, -1.270508, -2.636512, -0.805369, 1.570796, 2.018962],accel_mss,speed_ms,0,blend_radius_m)
  movel([0.454514, -1.271006, -2.636233, -0.805150, 1.570796, 2.025310],accel_mss,speed_ms,0,blend_radius_m)
  movel([0.460297, -1.271384, -2.636021, -0.804984, 1.570796, 2.031093],accel_mss,speed_ms,0,blend_radius_m)
  movel([0.464813, -1.271858, -2.635755, -0.804776, 1.570796, 2.035609],accel_mss,speed_ms,0,blend_radius_m)
  movel([0.475433, -1.273548, -2.634804, -0.804037, 1.570796, 2.046230],accel_mss,speed_ms,0,blend_radius_m)
  movel([0.480988, -1.274650, -2.634182, -0.803557, 1.570796, 2.051784],accel_mss,speed_ms,0,blend_radius_m)
  movel([0.485123, -1.275838, -2.633509, -0.803042, 1.570796, 2.055919],accel_mss,speed_ms,0,blend_radius_m)
  movel([0.486552, -1.276560, -2.633100, -0.802729, 1.570796, 2.057348],accel_mss,speed_ms,0,blend_radius_m)
  movel([0.487756, -1.277487, -2.632573, -0.802329, 1.570796, 2.058552],accel_mss,speed_ms,0,blend_radius_m)
  movel([0.489516, -1.279883, -2.631207, -0.801300, 1.570796, 2.060313],accel_mss,speed_ms,0,blend_radius_m)
  movel([0.490482, -1.282866, -2.629495, -0.800028, 1.570796, 2.061279],accel_mss,speed_ms,0,blend_radius_m)
  movel([0.490720, -1.286286, -2.627519, -0.798584, 1.570796, 2.061516],accel_mss,speed_ms,0,blend_radius_m)
  movel([0.490313, -1.289991, -2.625362, -0.797036, 1.570796, 2.061109],accel_mss,speed_ms,0,blend_radius_m)
  movel([0.489334, -1.293829, -2.623109, -0.795451, 1.570796, 2.060131],accel_mss,speed_ms,0,blend_radius_m)
  movel([0.487858, -1.297660, -2.620842, -0.793888, 1.570796, 2.058655],accel_mss,speed_ms,0,blend_radius_m)
  movel([0.485956, -1.301345, -2.618642, -0.792402, 1.570796, 2.056752],accel_mss,speed_ms,0,blend_radius_m)
  movel([0.483051, -1.305672, -2.616038, -0.790679, 1.570796, 2.053847],accel_mss,speed_ms,0,blend_radius_m)
  movel([0.481605, -1.307382, -2.615002, -0.790005, 1.570796, 2.052401],accel_mss,speed_ms,0,blend_radius_m)
  movel([0.480149, -1.308830, -2.614121, -0.789437, 1.570796, 2.050945],accel_mss,speed_ms,0,blend_radius_m)
  movel([0.478677, -1.310049, -2.613378, -0.788962, 1.570796, 2.049474],accel_mss,speed_ms,0,blend_radius_m)
  movel([0.477182, -1.311067, -2.612756, -0.788566, 1.570796, 2.047978],accel_mss,speed_ms,0,blend_radius_m)
  movel([0.474087, -1.312618, -2.611806, -0.787965, 1.570796, 2.044883],accel_mss,speed_ms,0,blend_radius_m)
  movel([0.470803, -1.313716, -2.611131, -0.787542, 1.570796, 2.041599],accel_mss,speed_ms,0,blend_radius_m)
  movel([0.467269, -1.314590, -2.610593, -0.787206, 1.570796, 2.038065],accel_mss,speed_ms,0,blend_radius_m)
  movel([0.459245, -1.316569, -2.609370, -0.786450, 1.570796, 2.030041],accel_mss,speed_ms,0,blend_radius_m)
  movel([0.458829, -1.316707, -2.609284, -0.786397, 1.570796, 2.029626],accel_mss,speed_ms,0,blend_radius_m)
  movel([0.458962, -1.316789, -2.609234, -0.786366, 1.570796, 2.029758],accel_mss,speed_ms,0,blend_radius_m)
  movel([0.460590, -1.316803, -2.609225, -0.786361, 1.570796, 2.031387],accel_mss,speed_ms,0,blend_radius_m)
  movel([0.467283, -1.316475, -2.609428, -0.786486, 1.570796, 2.038079],accel_mss,speed_ms,0,blend_radius_m)
  movel([0.478375, -1.315998, -2.609723, -0.786667, 1.570796, 2.049172],accel_mss,speed_ms,0,blend_radius_m)
  movel([0.471868, -1.319007, -2.607857, -0.785525, 1.570796, 2.042664],accel_mss,speed_ms,0,blend_radius_m)
  movel([0.464622, -1.322038, -2.605965, -0.784386, 1.570796, 2.035419],accel_mss,speed_ms,0,blend_radius_m)
  movel([0.456902, -1.325031, -2.604084, -0.783274, 1.570796, 2.027698],accel_mss,speed_ms,0,blend_radius_m)
  movel([0.448969, -1.327917, -2.602260, -0.782212, 1.570796, 2.019765],accel_mss,speed_ms,0,blend_radius_m)
  movel([0.433483, -1.333075, -2.598971, -0.780343, 1.570796, 2.004280],accel_mss,speed_ms,0,blend_radius_m)
  movel([0.426439, -1.335193, -2.597610, -0.779586, 1.570796, 1.997236],accel_mss,speed_ms,0,blend_radius_m)
  movel([0.420199, -1.336893, -2.596514, -0.778983, 1.570796, 1.990995],accel_mss,speed_ms,0,blend_radius_m)
  movel([0.411459, -1.342478, -2.592883, -0.777028, 1.570796, 1.982255],accel_mss,speed_ms,0,blend_radius_m)
  movel([0.402621, -1.348573, -2.588872, -0.774944, 1.570796, 1.973417],accel_mss,speed_ms,0,blend_radius_m)
  movel([0.384935, -1.361413, -2.580254, -0.770722, 1.570796, 1.955731],accel_mss,speed_ms,0,blend_radius_m)
  movel([0.376197, -1.367750, -2.575916, -0.768722, 1.570796, 1.946993],accel_mss,speed_ms,0,blend_radius_m)
  movel([0.367591, -1.373775, -2.571739, -0.766874, 1.570796, 1.938387],accel_mss,speed_ms,0,blend_radius_m)
  movel([0.359150, -1.379302, -2.567863, -0.765224, 1.570796, 1.929946],accel_mss,speed_ms,0,blend_radius_m)
  movel([0.350902, -1.384152, -2.564425, -0.763812, 1.570796, 1.921698],accel_mss,speed_ms,0,blend_radius_m)
  movel([0.347702, -1.385781, -2.563262, -0.763346, 1.570796, 1.918498],accel_mss,speed_ms,0,blend_radius_m)
  movel([0.344665, -1.387090, -2.562326, -0.762973, 1.570796, 1.915461],accel_mss,speed_ms,0,blend_radius_m)
  movel([0.341807, -1.388076, -2.561618, -0.762695, 1.570796, 1.912603],accel_mss,speed_ms,0,blend_radius_m)
  movel([0.339140, -1.388747, -2.561136, -0.762506, 1.570796, 1.909937],accel_mss,speed_ms,0,blend_radius_m)
  movel([0.336688, -1.389104, -2.560880, -0.762405, 1.570796, 1.907484],accel_mss,speed_ms,0,blend_radius_m)
  movel([0.334463, -1.389148, -2.560848, -0.762393, 1.570796, 1.905259],accel_mss,speed_ms,0,blend_radius_m)
  movel([0.332481, -1.388878, -2.561042, -0.762469, 1.570796, 1.903277],accel_mss,speed_ms,0,blend_radius_m)
  movel([0.330763, -1.388296, -2.561460, -0.762633, 1.570796, 1.901559],accel_mss,speed_ms,0,blend_radius_m)
  movel([0.329328, -1.387401, -2.562102, -0.762885, 1.570796, 1.900124],accel_mss,speed_ms,0,blend_radius_m)
  movel([0.328189, -1.386194, -2.562967, -0.763228, 1.570796, 1.898986],accel_mss,speed_ms,0,blend_radius_m)
  movel([0.327372, -1.384673, -2.564053, -0.763663, 1.570796, 1.898168],accel_mss,speed_ms,0,blend_radius_m)
  movel([0.326895, -1.382835, -2.565362, -0.764192, 1.570796, 1.897692],accel_mss,speed_ms,0,blend_radius_m)
  movel([0.326779, -1.380678, -2.566891, -0.764820, 1.570796, 1.897576],accel_mss,speed_ms,0,blend_radius_m)
  movel([0.327047, -1.378200, -2.568639, -0.765550, 1.570796, 1.897843],accel_mss,speed_ms,0,blend_radius_m)
  movel([0.327719, -1.375398, -2.570605, -0.766385, 1.570796, 1.898515],accel_mss,speed_ms,0,blend_radius_m)
  movel([0.328825, -1.372267, -2.572790, -0.767332, 1.570796, 1.899621],accel_mss,speed_ms,0,blend_radius_m)
  movel([0.331271, -1.373220, -2.572126, -0.767042, 1.570796, 1.902067],accel_mss,speed_ms,0,blend_radius_m)
  movel([0.332520, -1.373601, -2.571861, -0.766927, 1.570796, 1.903316],accel_mss,speed_ms,0,blend_radius_m)
  movel([0.333905, -1.373643, -2.571832, -0.766914, 1.570796, 1.904701],accel_mss,speed_ms,0,blend_radius_m)
  movel([0.335118, -1.373301, -2.572070, -0.767018, 1.570796, 1.905914],accel_mss,speed_ms,0,blend_radius_m)
  movel([0.336633, -1.372585, -2.572568, -0.767235, 1.570796, 1.907429],accel_mss,speed_ms,0,blend_radius_m)
  movel([0.340402, -1.370224, -2.574208, -0.767957, 1.570796, 1.911198],accel_mss,speed_ms,0,blend_radius_m)
  movel([0.344897, -1.366915, -2.576491, -0.768983, 1.570796, 1.915693],accel_mss,speed_ms,0,blend_radius_m)
  movel([0.349786, -1.363025, -2.579156, -0.770208, 1.570796, 1.920582],accel_mss,speed_ms,0,blend_radius_m)
  movel([0.359391, -1.354984, -2.584598, -0.772807, 1.570796, 1.930188],accel_mss,speed_ms,0,blend_radius_m)
  movel([0.366386, -1.349126, -2.588506, -0.774758, 1.570796, 1.937182],accel_mss,speed_ms,0,blend_radius_m)
  movel([0.372659, -1.344431, -2.591603, -0.776355, 1.570796, 1.943455],accel_mss,speed_ms,0,blend_radius_m)
  movel([0.378987, -1.339722, -2.594679, -0.777987, 1.570796, 1.949784],accel_mss,speed_ms,0,blend_radius_m)
  movel([0.366263, -1.342127, -2.593112, -0.777150, 1.570796, 1.937059],accel_mss,speed_ms,0,blend_radius_m)
  movel([0.359698, -1.343112, -2.592468, -0.776809, 1.570796, 1.930494],accel_mss,speed_ms,0,blend_radius_m)
  movel([0.353468, -1.343514, -2.592205, -0.776671, 1.570796, 1.924264],accel_mss,speed_ms,0,blend_radius_m)
  movel([0.350588, -1.343388, -2.592287, -0.776714, 1.570796, 1.921384],accel_mss,speed_ms,0,blend_radius_m)
  movel([0.347918, -1.342991, -2.592547, -0.776851, 1.570796, 1.918714],accel_mss,speed_ms,0,blend_radius_m)
  movel([0.345505, -1.342275, -2.593015, -0.777099, 1.570796, 1.916302],accel_mss,speed_ms,0,blend_radius_m)
  movel([0.343390, -1.341195, -2.593720, -0.777473, 1.570796, 1.914186],accel_mss,speed_ms,0,blend_radius_m)
  movel([0.341617, -1.339712, -2.594686, -0.777991, 1.570796, 1.912413],accel_mss,speed_ms,0,blend_radius_m)
  movel([0.340232, -1.337769, -2.595946, -0.778673, 1.570796, 1.911029],accel_mss,speed_ms,0,blend_radius_m)
  movel([0.339277, -1.335326, -2.597524, -0.779538, 1.570796, 1.910073],accel_mss,speed_ms,0,blend_radius_m)
  movel([0.338802, -1.332331, -2.599448, -0.780611, 1.570796, 1.909599],accel_mss,speed_ms,0,blend_radius_m)
  movel([0.338995, -1.328471, -2.601908, -0.782010, 1.570796, 1.909792],accel_mss,speed_ms,0,blend_radius_m)
  movel([0.340005, -1.324278, -2.604559, -0.783552, 1.570796, 1.910801],accel_mss,speed_ms,0,blend_radius_m)
  movel([0.341766, -1.319878, -2.607315, -0.785197, 1.570796, 1.912562],accel_mss,speed_ms,0,blend_radius_m)
  movel([0.344206, -1.315411, -2.610086, -0.786892, 1.570796, 1.915002],accel_mss,speed_ms,0,blend_radius_m)
  movel([0.347247, -1.311026, -2.612781, -0.788582, 1.570796, 1.918043],accel_mss,speed_ms,0,blend_radius_m)
  movel([0.350819, -1.306865, -2.615315, -0.790208, 1.570796, 1.921615],accel_mss,speed_ms,0,blend_radius_m)
  movel([0.354831, -1.303085, -2.617598, -0.791706, 1.570796, 1.925627],accel_mss,speed_ms,0,blend_radius_m)
  movel([0.359198, -1.299845, -2.619540, -0.793004, 1.570796, 1.929994],accel_mss,speed_ms,0,blend_radius_m)
  movel([0.361690, -1.298602, -2.620281, -0.793506, 1.570796, 1.932486],accel_mss,speed_ms,0,blend_radius_m)
  movel([0.364464, -1.297747, -2.620790, -0.793852, 1.570796, 1.935260],accel_mss,speed_ms,0,blend_radius_m)
  movel([0.366626, -1.297607, -2.620873, -0.793909, 1.570796, 1.937422],accel_mss,speed_ms,0,blend_radius_m)
  movel([0.367200, -1.297901, -2.620698, -0.793790, 1.570796, 1.937996],accel_mss,speed_ms,0,blend_radius_m)
  movel([0.367288, -1.298492, -2.620346, -0.793550, 1.570796, 1.938084],accel_mss,speed_ms,0,blend_radius_m)
  movel([0.365099, -1.299132, -2.619965, -0.793292, 1.570796, 1.935896],accel_mss,speed_ms,0,blend_radius_m)
  movel([0.363222, -1.299899, -2.619508, -0.792983, 1.570796, 1.934018],accel_mss,speed_ms,0,blend_radius_m)
  movel([0.361650, -1.300770, -2.618987, -0.792632, 1.570796, 1.932447],accel_mss,speed_ms,0,blend_radius_m)
  movel([0.360370, -1.301728, -2.618413, -0.792248, 1.570796, 1.931166],accel_mss,speed_ms,0,blend_radius_m)
  movel([0.359372, -1.302751, -2.617799, -0.791839, 1.570796, 1.930169],accel_mss,speed_ms,0,blend_radius_m)
  movel([0.358645, -1.303818, -2.617157, -0.791414, 1.570796, 1.929442],accel_mss,speed_ms,0,blend_radius_m)
  movel([0.358183, -1.304910, -2.616498, -0.790981, 1.570796, 1.928979],accel_mss,speed_ms,0,blend_radius_m)
  movel([0.357970, -1.306005, -2.615836, -0.790548, 1.570796, 1.928766],accel_mss,speed_ms,0,blend_radius_m)
  movel([0.358252, -1.308137, -2.614543, -0.789709, 1.570796, 1.929049],accel_mss,speed_ms,0,blend_radius_m)
  movel([0.359407, -1.310063, -2.613369, -0.788956, 1.570796, 1.930203],accel_mss,speed_ms,0,blend_radius_m)
  movel([0.361347, -1.311639, -2.612406, -0.788344, 1.570796, 1.932144],accel_mss,speed_ms,0,blend_radius_m)
  movel([0.363987, -1.312718, -2.611744, -0.787927, 1.570796, 1.934783],accel_mss,speed_ms,0,blend_radius_m)
  movel([0.365828, -1.313004, -2.611569, -0.787816, 1.570796, 1.936625],accel_mss,speed_ms,0,blend_radius_m)
  movel([0.368196, -1.313056, -2.611537, -0.787796, 1.570796, 1.938993],accel_mss,speed_ms,0,blend_radius_m)
  movel([0.374227, -1.312581, -2.611829, -0.787980, 1.570796, 1.945024],accel_mss,speed_ms,0,blend_radius_m)
  movel([0.381523, -1.311501, -2.612490, -0.788397, 1.570796, 1.952320],accel_mss,speed_ms,0,blend_radius_m)
  movel([0.389535, -1.310024, -2.613393, -0.788971, 1.570796, 1.960331],accel_mss,speed_ms,0,blend_radius_m)
  movel([0.405467, -1.306640, -2.615452, -0.790297, 1.570796, 1.976263],accel_mss,speed_ms,0,blend_radius_m)
  movel([0.417559, -1.303826, -2.617152, -0.791411, 1.570796, 1.988355],accel_mss,speed_ms,0,blend_radius_m)
  movel([0.423653, -1.302391, -2.618015, -0.791983, 1.570796, 1.994450],accel_mss,speed_ms,0,blend_radius_m)
  movel([0.426953, -1.301513, -2.618542, -0.792334, 1.570796, 1.997750],accel_mss,speed_ms,0,blend_radius_m)
  movel([0.429487, -1.300623, -2.619075, -0.792692, 1.570796, 2.000283],accel_mss,speed_ms,0,blend_radius_m)
  movel([0.430189, -1.300233, -2.619308, -0.792848, 1.570796, 2.000985],accel_mss,speed_ms,0,blend_radius_m)
  movel([0.430475, -1.299884, -2.619516, -0.792988, 1.570796, 2.001272],accel_mss,speed_ms,0,blend_radius_m)
  movel([0.430154, -1.299102, -2.619983, -0.793304, 1.570796, 2.000951],accel_mss,speed_ms,0,blend_radius_m)
  movel([0.428284, -1.297521, -2.620924, -0.793944, 1.570796, 1.999081],accel_mss,speed_ms,0,blend_radius_m)
  movel([0.425890, -1.296368, -2.621608, -0.794413, 1.570796, 1.996686],accel_mss,speed_ms,0,blend_radius_m)
  movel([0.420503, -1.294187, -2.622898, -0.795304, 1.570796, 1.991299],accel_mss,speed_ms,0,blend_radius_m)
  movel([0.418003, -1.292571, -2.623850, -0.795968, 1.570796, 1.988799],accel_mss,speed_ms,0,blend_radius_m)
  movel([0.415957, -1.290209, -2.625235, -0.796946, 1.570796, 1.986753],accel_mss,speed_ms,0,blend_radius_m)
  movel([0.415181, -1.288649, -2.626145, -0.797594, 1.570796, 1.985977],accel_mss,speed_ms,0,blend_radius_m)
  movel([0.414610, -1.286789, -2.627228, -0.798373, 1.570796, 1.985406],accel_mss,speed_ms,0,blend_radius_m)
  movel([0.414281, -1.284581, -2.628506, -0.799302, 1.570796, 1.985077],accel_mss,speed_ms,0,blend_radius_m)
  movel([0.414220, -1.281988, -2.630000, -0.800401, 1.570796, 1.985016],accel_mss,speed_ms,0,blend_radius_m)
  movel([0.414685, -1.278356, -2.632078, -0.801955, 1.570796, 1.985482],accel_mss,speed_ms,0,blend_radius_m)
  movel([0.415805, -1.274724, -2.634140, -0.803525, 1.570796, 1.986602],accel_mss,speed_ms,0,blend_radius_m)
  movel([0.417510, -1.271103, -2.636179, -0.805107, 1.570796, 1.988307],accel_mss,speed_ms,0,blend_radius_m)
  movel([0.419716, -1.267508, -2.638187, -0.806694, 1.570796, 1.990513],accel_mss,speed_ms,0,blend_radius_m)
  movel([0.422352, -1.263951, -2.640159, -0.808279, 1.570796, 1.993149],accel_mss,speed_ms,0,blend_radius_m)
  movel([0.425336, -1.260449, -2.642085, -0.809855, 1.570796, 1.996132],accel_mss,speed_ms,0,blend_radius_m)
  movel([0.428586, -1.257023, -2.643955, -0.811411, 1.570796, 1.999383],accel_mss,speed_ms,0,blend_radius_m)
  movel([0.432023, -1.253682, -2.645764, -0.812942, 1.570796, 2.002819],accel_mss,speed_ms,0,blend_radius_m)
  movel([0.438800, -1.247807, -2.648915, -0.815668, 1.570796, 2.009596],accel_mss,speed_ms,0,blend_radius_m)
  movel([0.445021, -1.243212, -2.651349, -0.817828, 1.570796, 2.015818],accel_mss,speed_ms,0,blend_radius_m)
  movel([0.450384, -1.239833, -2.653124, -0.819432, 1.570796, 2.021180],accel_mss,speed_ms,0,blend_radius_m)
  movel([0.454585, -1.237590, -2.654295, -0.820505, 1.570796, 2.025381],accel_mss,speed_ms,0,blend_radius_m)
  movel([0.460811, -1.234970, -2.655654, -0.821764, 1.570796, 2.031608],accel_mss,speed_ms,0,blend_radius_m)
  movel([0.466812, -1.233235, -2.656550, -0.822603, 1.570796, 2.037608],accel_mss,speed_ms,0,blend_radius_m)
  movel([0.472511, -1.232358, -2.657002, -0.823029, 1.570796, 2.043308],accel_mss,speed_ms,0,blend_radius_m)
  movel([0.477835, -1.232322, -2.657021, -0.823046, 1.570796, 2.048631],accel_mss,speed_ms,0,blend_radius_m)
  movel([0.482714, -1.233091, -2.656625, -0.822673, 1.570796, 2.053511],accel_mss,speed_ms,0,blend_radius_m)
  movel([0.487084, -1.234638, -2.655826, -0.821925, 1.570796, 2.057881],accel_mss,speed_ms,0,blend_radius_m)
  movel([0.490883, -1.236920, -2.654643, -0.820826, 1.570796, 2.061679],accel_mss,speed_ms,0,blend_radius_m)
  movel([0.494051, -1.239897, -2.653091, -0.819402, 1.570796, 2.064847],accel_mss,speed_ms,0,blend_radius_m)
  movel([0.496320, -1.243132, -2.651391, -0.817865, 1.570796, 2.067116],accel_mss,speed_ms,0,blend_radius_m)
  movel([0.498191, -1.246657, -2.649526, -0.816206, 1.570796, 2.068987],accel_mss,speed_ms,0,blend_radius_m)
  movel([0.499961, -1.250174, -2.647651, -0.814565, 1.570796, 2.070757],accel_mss,speed_ms,0,blend_radius_m)
  movel([0.501923, -1.253391, -2.645921, -0.813076, 1.570796, 2.072720],accel_mss,speed_ms,0,blend_radius_m)
  movel([0.504362, -1.256038, -2.644490, -0.811861, 1.570796, 2.075158],accel_mss,speed_ms,0,blend_radius_m)
  movel([0.505848, -1.257060, -2.643934, -0.811394, 1.570796, 2.076644],accel_mss,speed_ms,0,blend_radius_m)
  movel([0.507562, -1.257835, -2.643513, -0.811041, 1.570796, 2.078358],accel_mss,speed_ms,0,blend_radius_m)
  movel([0.509541, -1.258331, -2.643243, -0.810815, 1.570796, 2.080338],accel_mss,speed_ms,0,blend_radius_m)
  movel([0.511819, -1.258515, -2.643142, -0.810732, 1.570796, 2.082615],accel_mss,speed_ms,0,blend_radius_m)
  movel([0.514435, -1.258350, -2.643232, -0.810807, 1.570796, 2.085231],accel_mss,speed_ms,0,blend_radius_m)
  movel([0.517427, -1.257806, -2.643529, -0.811054, 1.570796, 2.088223],accel_mss,speed_ms,0,blend_radius_m)
  movel([0.520140, -1.256933, -2.644004, -0.811452, 1.570796, 2.090936],accel_mss,speed_ms,0,blend_radius_m)
  movel([0.522509, -1.255711, -2.644667, -0.812011, 1.570796, 2.093306],accel_mss,speed_ms,0,blend_radius_m)
  movel([0.524533, -1.254206, -2.645482, -0.812701, 1.570796, 2.095329],accel_mss,speed_ms,0,blend_radius_m)
  movel([0.526215, -1.252490, -2.646407, -0.813492, 1.570796, 2.097011],accel_mss,speed_ms,0,blend_radius_m)
  movel([0.527545, -1.250637, -2.647402, -0.814350, 1.570796, 2.098342],accel_mss,speed_ms,0,blend_radius_m)
  movel([0.528526, -1.248712, -2.648432, -0.815245, 1.570796, 2.099322],accel_mss,speed_ms,0,blend_radius_m)
  movel([0.529151, -1.246798, -2.649451, -0.816140, 1.570796, 2.099947],accel_mss,speed_ms,0,blend_radius_m)
  movel([0.529414, -1.244964, -2.650424, -0.817001, 1.570796, 2.100210],accel_mss,speed_ms,0,blend_radius_m)
  movel([0.529313, -1.243286, -2.651310, -0.817793, 1.570796, 2.100109],accel_mss,speed_ms,0,blend_radius_m)
  movel([0.528840, -1.241846, -2.652068, -0.818474, 1.570796, 2.099637],accel_mss,speed_ms,0,blend_radius_m)
  movel([0.527989, -1.240723, -2.652658, -0.819008, 1.570796, 2.098786],accel_mss,speed_ms,0,blend_radius_m)
  movel([0.526761, -1.239990, -2.653042, -0.819357, 1.570796, 2.097558],accel_mss,speed_ms,0,blend_radius_m)
  movel([0.525154, -1.239726, -2.653180, -0.819483, 1.570796, 2.095950],accel_mss,speed_ms,0,blend_radius_m)
  movel([0.523162, -1.240011, -2.653031, -0.819347, 1.570796, 2.093958],accel_mss,speed_ms,0,blend_radius_m)
  movel([0.520787, -1.240918, -2.652556, -0.818915, 1.570796, 2.091583],accel_mss,speed_ms,0,blend_radius_m)
  movel([0.518035, -1.242521, -2.651713, -0.818155, 1.570796, 2.088831],accel_mss,speed_ms,0,blend_radius_m)
  movel([0.519548, -1.242789, -2.651572, -0.818028, 1.570796, 2.090344],accel_mss,speed_ms,0,blend_radius_m)
  movel([0.520623, -1.243354, -2.651274, -0.817760, 1.570796, 2.091420],accel_mss,speed_ms,0,blend_radius_m)
  movel([0.521253, -1.244166, -2.650846, -0.817377, 1.570796, 2.092050],accel_mss,speed_ms,0,blend_radius_m)
  movel([0.521427, -1.245188, -2.650305, -0.816896, 1.570796, 2.092223],accel_mss,speed_ms,0,blend_radius_m)
  movel([0.521141, -1.246373, -2.649677, -0.816339, 1.570796, 2.091938],accel_mss,speed_ms,0,blend_radius_m)
  movel([0.520392, -1.247681, -2.648982, -0.815727, 1.570796, 2.091188],accel_mss,speed_ms,0,blend_radius_m)
  movel([0.519169, -1.249068, -2.648242, -0.815079, 1.570796, 2.089966],accel_mss,speed_ms,0,blend_radius_m)
  movel([0.517466, -1.250495, -2.647478, -0.814415, 1.570796, 2.088263],accel_mss,speed_ms,0,blend_radius_m)
  movel([0.514332, -1.252431, -2.646439, -0.813519, 1.570796, 2.085129],accel_mss,speed_ms,0,blend_radius_m)
  movel([0.511473, -1.253485, -2.645871, -0.813033, 1.570796, 2.082269],accel_mss,speed_ms,0,blend_radius_m)
  movel([0.508906, -1.253742, -2.645732, -0.812915, 1.570796, 2.079702],accel_mss,speed_ms,0,blend_radius_m)
  movel([0.506657, -1.253290, -2.645976, -0.813123, 1.570796, 2.077454],accel_mss,speed_ms,0,blend_radius_m)
  movel([0.504753, -1.252207, -2.646559, -0.813623, 1.570796, 2.075549],accel_mss,speed_ms,0,blend_radius_m)
  movel([0.503219, -1.250573, -2.647436, -0.814379, 1.570796, 2.074015],accel_mss,speed_ms,0,blend_radius_m)
  movel([0.502087, -1.248468, -2.648562, -0.815359, 1.570796, 2.072883],accel_mss,speed_ms,0,blend_radius_m)
  movel([0.501387, -1.245964, -2.649894, -0.816531, 1.570796, 2.072183],accel_mss,speed_ms,0,blend_radius_m)
  movel([0.501156, -1.243138, -2.651388, -0.817863, 1.570796, 2.071952],accel_mss,speed_ms,0,blend_radius_m)
  movel([0.501425, -1.240070, -2.653000, -0.819319, 1.570796, 2.072221],accel_mss,speed_ms,0,blend_radius_m)
  movel([0.502231, -1.236839, -2.654685, -0.820865, 1.570796, 2.073027],accel_mss,speed_ms,0,blend_radius_m)
  movel([0.503615, -1.233519, -2.656404, -0.822466, 1.570796, 2.074412],accel_mss,speed_ms,0,blend_radius_m)
  movel([0.505607, -1.230200, -2.658110, -0.824079, 1.570796, 2.076403],accel_mss,speed_ms,0,blend_radius_m)
  movel([0.508244, -1.226968, -2.659758, -0.825663, 1.570796, 2.079040],accel_mss,speed_ms,0,blend_radius_m)
  movel([0.511562, -1.223907, -2.661309, -0.827173, 1.570796, 2.082359],accel_mss,speed_ms,0,blend_radius_m)
  movel([0.515588, -1.221116, -2.662713, -0.828560, 1.570796, 2.086385],accel_mss,speed_ms,0,blend_radius_m)
  movel([0.518604, -1.219449, -2.663547, -0.829393, 1.570796, 2.089400],accel_mss,speed_ms,0,blend_radius_m)
  movel([0.521611, -1.218042, -2.664249, -0.830098, 1.570796, 2.092408],accel_mss,speed_ms,0,blend_radius_m)
  movel([0.524583, -1.216906, -2.664814, -0.830669, 1.570796, 2.095380],accel_mss,speed_ms,0,blend_radius_m)
  movel([0.527498, -1.216043, -2.665243, -0.831103, 1.570796, 2.098295],accel_mss,speed_ms,0,blend_radius_m)
  movel([0.530329, -1.215456, -2.665534, -0.831400, 1.570796, 2.101125],accel_mss,speed_ms,0,blend_radius_m)
  movel([0.533049, -1.215154, -2.665683, -0.831552, 1.570796, 2.103845],accel_mss,speed_ms,0,blend_radius_m)
  movel([0.535632, -1.215139, -2.665690, -0.831559, 1.570796, 2.106428],accel_mss,speed_ms,0,blend_radius_m)
  movel([0.538053, -1.215414, -2.665554, -0.831421, 1.570796, 2.108849],accel_mss,speed_ms,0,blend_radius_m)
  movel([0.540290, -1.215980, -2.665274, -0.831135, 1.570796, 2.111086],accel_mss,speed_ms,0,blend_radius_m)
  movel([0.542318, -1.216837, -2.664849, -0.830703, 1.570796, 2.113114],accel_mss,speed_ms,0,blend_radius_m)
  movel([0.544112, -1.217990, -2.664275, -0.830124, 1.570796, 2.114908],accel_mss,speed_ms,0,blend_radius_m)
  movel([0.545650, -1.219436, -2.663554, -0.829399, 1.570796, 2.116446],accel_mss,speed_ms,0,blend_radius_m)
  movel([0.546907, -1.221177, -2.662683, -0.828530, 1.570796, 2.117703],accel_mss,speed_ms,0,blend_radius_m)
  movel([0.547866, -1.223209, -2.661661, -0.827519, 1.570796, 2.118662],accel_mss,speed_ms,0,blend_radius_m)
  movel([0.548503, -1.225534, -2.660486, -0.826369, 1.570796, 2.119300],accel_mss,speed_ms,0,blend_radius_m)
  movel([0.548798, -1.228149, -2.659157, -0.825083, 1.570796, 2.119594],accel_mss,speed_ms,0,blend_radius_m)
  movel([0.548394, -1.231056, -2.657671, -0.823662, 1.570796, 2.119191],accel_mss,speed_ms,0,blend_radius_m)
  movel([0.547374, -1.234387, -2.655956, -0.822046, 1.570796, 2.118170],accel_mss,speed_ms,0,blend_radius_m)
  movel([0.546349, -1.237281, -2.654455, -0.820653, 1.570796, 2.117145],accel_mss,speed_ms,0,blend_radius_m)
  movel([0.545903, -1.238901, -2.653611, -0.819877, 1.570796, 2.116699],accel_mss,speed_ms,0,blend_radius_m)
  movel([0.546549, -1.239688, -2.653200, -0.819501, 1.570796, 2.117346],accel_mss,speed_ms,0,blend_radius_m)
  movel([0.547986, -1.240608, -2.652718, -0.819063, 1.570796, 2.118783],accel_mss,speed_ms,0,blend_radius_m)
  movel([0.549570, -1.241621, -2.652186, -0.818581, 1.570796, 2.120367],accel_mss,speed_ms,0,blend_radius_m)
  movel([0.550668, -1.242681, -2.651629, -0.818079, 1.570796, 2.121464],accel_mss,speed_ms,0,blend_radius_m)
  movel([0.551522, -1.244564, -2.650636, -0.817190, 1.570796, 2.122318],accel_mss,speed_ms,0,blend_radius_m)
  movel([0.551940, -1.246581, -2.649566, -0.816241, 1.570796, 2.122736],accel_mss,speed_ms,0,blend_radius_m)
  movel([0.551953, -1.248705, -2.648436, -0.815248, 1.570796, 2.122750],accel_mss,speed_ms,0,blend_radius_m)
  movel([0.551593, -1.250900, -2.647261, -0.814228, 1.570796, 2.122389],accel_mss,speed_ms,0,blend_radius_m)
  movel([0.550886, -1.253137, -2.646059, -0.813194, 1.570796, 2.121682],accel_mss,speed_ms,0,blend_radius_m)
  movel([0.549872, -1.255378, -2.644848, -0.812164, 1.570796, 2.120668],accel_mss,speed_ms,0,blend_radius_m)
  movel([0.548573, -1.257598, -2.643642, -0.811149, 1.570796, 2.119370],accel_mss,speed_ms,0,blend_radius_m)
  movel([0.547025, -1.259767, -2.642458, -0.810164, 1.570796, 2.117821],accel_mss,speed_ms,0,blend_radius_m)
  movel([0.545252, -1.261856, -2.641313, -0.809220, 1.570796, 2.116048],accel_mss,speed_ms,0,blend_radius_m)
  movel([0.543286, -1.263834, -2.640223, -0.808331, 1.570796, 2.114082],accel_mss,speed_ms,0,blend_radius_m)
  movel([0.541155, -1.265675, -2.639205, -0.807509, 1.570796, 2.111951],accel_mss,speed_ms,0,blend_radius_m)
  speed_ms = 0.003
  movel([0.541155, -1.258681, -2.635807, -0.817901, 1.570796, 2.111951],accel_mss,speed_ms,0,blend_radius_m)
  speed_ms = 0.1
  movel([0.541155, -1.231973, -2.621944, -0.858472, 1.570796, 2.111951],accel_mss,speed_ms,0,blend_radius_m)
  #M_RunCode9
  movel([0.555888, -1.230851, -2.622537, -0.859001, 1.570796, 2.126684],accel_mss,speed_ms,0,blend_radius_m)
  #M_RunCode3
  movel([0.555888, -1.257572, -2.636415, -0.818402, 1.570796, 2.126684],accel_mss,speed_ms,0,blend_radius_m)
  speed_ms = 0.003
  movel([0.555888, -1.264570, -2.639817, -0.808002, 1.570796, 2.126684],accel_mss,speed_ms,0,blend_radius_m)
  speed_ms = 0.007
  movel([0.556708, -1.262696, -2.640851, -0.808842, 1.570796, 2.127505],accel_mss,speed_ms,0,blend_radius_m)
  movel([0.558883, -1.258875, -2.642946, -0.810568, 1.570796, 2.129679],accel_mss,speed_ms,0,blend_radius_m)
  movel([0.560835, -1.255136, -2.644978, -0.812274, 1.570796, 2.131631],accel_mss,speed_ms,0,blend_radius_m)
  movel([0.561371, -1.253369, -2.645933, -0.813087, 1.570796, 2.132167],accel_mss,speed_ms,0,blend_radius_m)
  movel([0.561424, -1.251703, -2.646830, -0.813856, 1.570796, 2.132220],accel_mss,speed_ms,0,blend_radius_m)
  movel([0.561823, -1.252697, -2.646295, -0.813396, 1.570796, 2.132619],accel_mss,speed_ms,0,blend_radius_m)
  movel([0.562077, -1.254762, -2.645181, -0.812446, 1.570796, 2.132873],accel_mss,speed_ms,0,blend_radius_m)
  movel([0.561745, -1.256887, -2.644029, -0.811473, 1.570796, 2.132541],accel_mss,speed_ms,0,blend_radius_m)
  movel([0.561009, -1.259053, -2.642849, -0.810487, 1.570796, 2.131805],accel_mss,speed_ms,0,blend_radius_m)
  movel([0.560050, -1.261245, -2.641649, -0.809496, 1.570796, 2.130847],accel_mss,speed_ms,0,blend_radius_m)
  movel([0.558184, -1.265634, -2.639228, -0.807527, 1.570796, 2.128981],accel_mss,speed_ms,0,blend_radius_m)
  movel([0.557629, -1.267804, -2.638023, -0.806563, 1.570796, 2.128425],accel_mss,speed_ms,0,blend_radius_m)
  movel([0.557564, -1.269935, -2.636833, -0.805621, 1.570796, 2.128360],accel_mss,speed_ms,0,blend_radius_m)
  movel([0.558013, -1.272106, -2.635616, -0.804667, 1.570796, 2.128809],accel_mss,speed_ms,0,blend_radius_m)
  movel([0.558382, -1.273196, -2.635002, -0.804191, 1.570796, 2.129178],accel_mss,speed_ms,0,blend_radius_m)
  movel([0.558780, -1.273706, -2.634715, -0.803968, 1.570796, 2.129576],accel_mss,speed_ms,0,blend_radius_m)
  movel([0.560056, -1.273237, -2.634979, -0.804173, 1.570796, 2.130853],accel_mss,speed_ms,0,blend_radius_m)
  movel([0.561102, -1.272903, -2.635167, -0.804319, 1.570796, 2.131898],accel_mss,speed_ms,0,blend_radius_m)
  movel([0.562138, -1.272761, -2.635247, -0.804381, 1.570796, 2.132934],accel_mss,speed_ms,0,blend_radius_m)
  movel([0.563992, -1.272958, -2.635136, -0.804295, 1.570796, 2.134788],accel_mss,speed_ms,0,blend_radius_m)
  movel([0.565214, -1.273424, -2.634874, -0.804091, 1.570796, 2.136011],accel_mss,speed_ms,0,blend_radius_m)
  movel([0.565941, -1.274124, -2.634479, -0.803786, 1.570796, 2.136738],accel_mss,speed_ms,0,blend_radius_m)
  movel([0.566309, -1.275019, -2.633973, -0.803397, 1.570796, 2.137105],accel_mss,speed_ms,0,blend_radius_m)
  movel([0.566515, -1.277260, -2.632702, -0.802427, 1.570796, 2.137311],accel_mss,speed_ms,0,blend_radius_m)
  movel([0.566924, -1.279873, -2.631212, -0.801304, 1.570796, 2.137721],accel_mss,speed_ms,0,blend_radius_m)
  movel([0.568152, -1.283006, -2.629414, -0.799968, 1.570796, 2.138949],accel_mss,speed_ms,0,blend_radius_m)
  movel([0.569521, -1.286022, -2.627672, -0.798694, 1.570796, 2.140318],accel_mss,speed_ms,0,blend_radius_m)
  movel([0.570695, -1.289145, -2.625856, -0.797388, 1.570796, 2.141492],accel_mss,speed_ms,0,blend_radius_m)
  movel([0.571345, -1.292588, -2.623840, -0.795961, 1.570796, 2.142141],accel_mss,speed_ms,0,blend_radius_m)
  movel([0.571345, -1.294616, -2.622645, -0.795128, 1.570796, 2.142141],accel_mss,speed_ms,0,blend_radius_m)
  movel([0.571088, -1.296726, -2.621396, -0.794267, 1.570796, 2.141884],accel_mss,speed_ms,0,blend_radius_m)
  movel([0.570075, -1.301077, -2.618803, -0.792509, 1.570796, 2.140871],accel_mss,speed_ms,0,blend_radius_m)
  movel([0.568812, -1.305418, -2.616191, -0.790780, 1.570796, 2.139608],accel_mss,speed_ms,0,blend_radius_m)
  movel([0.567799, -1.309540, -2.613689, -0.789160, 1.570796, 2.138595],accel_mss,speed_ms,0,blend_radius_m)
  movel([0.566993, -1.316103, -2.609658, -0.786627, 1.570796, 2.137789],accel_mss,speed_ms,0,blend_radius_m)
  movel([0.566727, -1.318878, -2.607937, -0.785574, 1.570796, 2.137523],accel_mss,speed_ms,0,blend_radius_m)
  movel([0.566292, -1.321541, -2.606276, -0.784572, 1.570796, 2.137088],accel_mss,speed_ms,0,blend_radius_m)
  movel([0.565492, -1.324262, -2.604569, -0.783559, 1.570796, 2.136289],accel_mss,speed_ms,0,blend_radius_m)
  movel([0.564136, -1.327201, -2.602713, -0.782474, 1.570796, 2.134933],accel_mss,speed_ms,0,blend_radius_m)
  movel([0.562034, -1.330522, -2.600603, -0.781264, 1.570796, 2.132830],accel_mss,speed_ms,0,blend_radius_m)
  movel([0.559007, -1.334381, -2.598133, -0.779876, 1.570796, 2.129803],accel_mss,speed_ms,0,blend_radius_m)
  movel([0.556276, -1.337375, -2.596201, -0.778812, 1.570796, 2.127072],accel_mss,speed_ms,0,blend_radius_m)
  movel([0.553547, -1.339954, -2.594528, -0.777906, 1.570796, 2.124343],accel_mss,speed_ms,0,blend_radius_m)
  movel([0.550819, -1.342145, -2.593101, -0.777144, 1.570796, 2.121615],accel_mss,speed_ms,0,blend_radius_m)
  movel([0.548098, -1.343971, -2.591905, -0.776513, 1.570796, 2.118894],accel_mss,speed_ms,0,blend_radius_m)
  movel([0.545381, -1.345457, -2.590929, -0.776003, 1.570796, 2.116178],accel_mss,speed_ms,0,blend_radius_m)
  movel([0.542679, -1.346622, -2.590161, -0.775606, 1.570796, 2.113476],accel_mss,speed_ms,0,blend_radius_m)
  movel([0.539994, -1.347491, -2.589588, -0.775311, 1.570796, 2.110790],accel_mss,speed_ms,0,blend_radius_m)
  movel([0.537330, -1.348080, -2.589198, -0.775111, 1.570796, 2.108126],accel_mss,speed_ms,0,blend_radius_m)
  movel([0.534688, -1.348416, -2.588976, -0.774997, 1.570796, 2.105485],accel_mss,speed_ms,0,blend_radius_m)
  movel([0.532078, -1.348512, -2.588912, -0.774965, 1.570796, 2.102874],accel_mss,speed_ms,0,blend_radius_m)
  movel([0.526970, -1.348073, -2.589203, -0.775113, 1.570796, 2.097767],accel_mss,speed_ms,0,blend_radius_m)
  movel([0.522049, -1.346913, -2.589969, -0.775507, 1.570796, 2.092845],accel_mss,speed_ms,0,blend_radius_m)
  movel([0.517368, -1.345175, -2.591114, -0.776100, 1.570796, 2.088164],accel_mss,speed_ms,0,blend_radius_m)
  movel([0.513292, -1.343080, -2.592489, -0.776820, 1.570796, 2.084089],accel_mss,speed_ms,0,blend_radius_m)
  movel([0.508143, -1.340288, -2.594311, -0.777790, 1.570796, 2.078939],accel_mss,speed_ms,0,blend_radius_m)
  movel([0.502147, -1.337535, -2.596098, -0.778756, 1.570796, 2.072944],accel_mss,speed_ms,0,blend_radius_m)
  movel([0.498911, -1.336404, -2.596829, -0.779156, 1.570796, 2.069707],accel_mss,speed_ms,0,blend_radius_m)
  movel([0.495562, -1.335556, -2.597376, -0.779457, 1.570796, 2.066358],accel_mss,speed_ms,0,blend_radius_m)
  movel([0.492137, -1.335084, -2.597680, -0.779625, 1.570796, 2.062933],accel_mss,speed_ms,0,blend_radius_m)
  movel([0.488671, -1.335076, -2.597685, -0.779628, 1.570796, 2.059468],accel_mss,speed_ms,0,blend_radius_m)
  movel([0.485210, -1.335617, -2.597337, -0.779435, 1.570796, 2.056006],accel_mss,speed_ms,0,blend_radius_m)
  movel([0.481794, -1.336792, -2.596579, -0.779018, 1.570796, 2.052590],accel_mss,speed_ms,0,blend_radius_m)
  movel([0.480116, -1.337641, -2.596029, -0.778718, 1.570796, 2.050912],accel_mss,speed_ms,0,blend_radius_m)
  movel([0.478464, -1.338681, -2.595356, -0.778352, 1.570796, 2.049260],accel_mss,speed_ms,0,blend_radius_m)
  movel([0.476846, -1.339918, -2.594552, -0.777919, 1.570796, 2.047643],accel_mss,speed_ms,0,blend_radius_m)
  movel([0.475267, -1.341363, -2.593611, -0.777415, 1.570796, 2.046063],accel_mss,speed_ms,0,blend_radius_m)
  movel([0.473729, -1.343026, -2.592524, -0.776839, 1.570796, 2.044526],accel_mss,speed_ms,0,blend_radius_m)
  movel([0.472245, -1.344912, -2.591287, -0.776190, 1.570796, 2.043041],accel_mss,speed_ms,0,blend_radius_m)
  movel([0.469443, -1.349395, -2.588327, -0.774667, 1.570796, 2.040239],accel_mss,speed_ms,0,blend_radius_m)
  movel([0.468650, -1.351589, -2.586868, -0.773932, 1.570796, 2.039446],accel_mss,speed_ms,0,blend_radius_m)
  movel([0.468274, -1.353775, -2.585408, -0.773206, 1.570796, 2.039070],accel_mss,speed_ms,0,blend_radius_m)
  movel([0.468350, -1.355927, -2.583964, -0.772498, 1.570796, 2.039147],accel_mss,speed_ms,0,blend_radius_m)
  movel([0.468904, -1.358023, -2.582552, -0.771814, 1.570796, 2.039701],accel_mss,speed_ms,0,blend_radius_m)
  movel([0.471289, -1.355291, -2.584392, -0.772706, 1.570796, 2.042085],accel_mss,speed_ms,0,blend_radius_m)
  movel([0.473831, -1.352788, -2.586068, -0.773533, 1.570796, 2.044627],accel_mss,speed_ms,0,blend_radius_m)
  movel([0.476502, -1.350530, -2.587573, -0.774286, 1.570796, 2.047299],accel_mss,speed_ms,0,blend_radius_m)
  movel([0.479279, -1.348525, -2.588904, -0.774960, 1.570796, 2.050075],accel_mss,speed_ms,0,blend_radius_m)
  movel([0.482131, -1.346786, -2.590053, -0.775550, 1.570796, 2.052927],accel_mss,speed_ms,0,blend_radius_m)
  movel([0.485028, -1.345321, -2.591019, -0.776050, 1.570796, 2.055824],accel_mss,speed_ms,0,blend_radius_m)
  movel([0.487945, -1.344138, -2.591796, -0.776456, 1.570796, 2.058741],accel_mss,speed_ms,0,blend_radius_m)
  movel([0.490851, -1.343251, -2.592377, -0.776761, 1.570796, 2.061647],accel_mss,speed_ms,0,blend_radius_m)
  movel([0.493716, -1.342668, -2.592759, -0.776963, 1.570796, 2.064513],accel_mss,speed_ms,0,blend_radius_m)
  movel([0.496514, -1.342393, -2.592938, -0.777058, 1.570796, 2.067311],accel_mss,speed_ms,0,blend_radius_m)
  movel([0.499215, -1.342436, -2.592910, -0.777043, 1.570796, 2.070012],accel_mss,speed_ms,0,blend_radius_m)
  movel([0.501789, -1.342804, -2.592669, -0.776915, 1.570796, 2.072586],accel_mss,speed_ms,0,blend_radius_m)
  movel([0.504209, -1.343504, -2.592211, -0.776674, 1.570796, 2.075005],accel_mss,speed_ms,0,blend_radius_m)
  movel([0.506448, -1.344538, -2.591533, -0.776318, 1.570796, 2.077245],accel_mss,speed_ms,0,blend_radius_m)
  movel([0.508478, -1.345913, -2.590628, -0.775847, 1.570796, 2.079274],accel_mss,speed_ms,0,blend_radius_m)
  movel([0.510273, -1.347632, -2.589494, -0.775263, 1.570796, 2.081069],accel_mss,speed_ms,0,blend_radius_m)
  movel([0.511513, -1.349263, -2.588415, -0.774711, 1.570796, 2.082309],accel_mss,speed_ms,0,blend_radius_m)
  movel([0.512476, -1.351015, -2.587251, -0.774124, 1.570796, 2.083272],accel_mss,speed_ms,0,blend_radius_m)
  movel([0.513179, -1.352870, -2.586014, -0.773506, 1.570796, 2.083975],accel_mss,speed_ms,0,blend_radius_m)
  movel([0.513634, -1.354812, -2.584713, -0.772864, 1.570796, 2.084430],accel_mss,speed_ms,0,blend_radius_m)
  movel([0.513841, -1.358895, -2.581962, -0.771531, 1.570796, 2.084637],accel_mss,speed_ms,0,blend_radius_m)
  movel([0.513196, -1.363144, -2.579075, -0.770170, 1.570796, 2.083992],accel_mss,speed_ms,0,blend_radius_m)
  movel([0.511798, -1.367440, -2.576130, -0.768819, 1.570796, 2.082594],accel_mss,speed_ms,0,blend_radius_m)
  movel([0.509737, -1.371671, -2.573204, -0.767514, 1.570796, 2.080533],accel_mss,speed_ms,0,blend_radius_m)
  movel([0.507105, -1.375728, -2.570375, -0.766286, 1.570796, 2.077901],accel_mss,speed_ms,0,blend_radius_m)
  movel([0.503989, -1.379510, -2.567716, -0.765163, 1.570796, 2.074786],accel_mss,speed_ms,0,blend_radius_m)
  movel([0.500471, -1.382916, -2.565304, -0.764169, 1.570796, 2.071268],accel_mss,speed_ms,0,blend_radius_m)
  movel([0.496631, -1.385844, -2.563217, -0.763328, 1.570796, 2.067428],accel_mss,speed_ms,0,blend_radius_m)
  movel([0.492546, -1.388200, -2.561529, -0.762660, 1.570796, 2.063343],accel_mss,speed_ms,0,blend_radius_m)
  movel([0.490432, -1.389133, -2.560859, -0.762397, 1.570796, 2.061228],accel_mss,speed_ms,0,blend_radius_m)
  movel([0.488284, -1.389888, -2.560315, -0.762186, 1.570796, 2.059080],accel_mss,speed_ms,0,blend_radius_m)
  movel([0.486107, -1.390450, -2.559910, -0.762029, 1.570796, 2.056903],accel_mss,speed_ms,0,blend_radius_m)
  movel([0.483914, -1.390810, -2.559650, -0.761929, 1.570796, 2.054710],accel_mss,speed_ms,0,blend_radius_m)
  movel([0.481710, -1.390951, -2.559548, -0.761890, 1.570796, 2.052506],accel_mss,speed_ms,0,blend_radius_m)
  movel([0.479505, -1.390865, -2.559610, -0.761914, 1.570796, 2.050301],accel_mss,speed_ms,0,blend_radius_m)
  movel([0.477302, -1.390538, -2.559846, -0.762005, 1.570796, 2.048099],accel_mss,speed_ms,0,blend_radius_m)
  movel([0.475117, -1.389954, -2.560267, -0.762167, 1.570796, 2.045914],accel_mss,speed_ms,0,blend_radius_m)
  movel([0.472951, -1.389103, -2.560880, -0.762406, 1.570796, 2.043748],accel_mss,speed_ms,0,blend_radius_m)
  movel([0.470815, -1.387971, -2.561694, -0.762724, 1.570796, 2.041612],accel_mss,speed_ms,0,blend_radius_m)
  movel([0.469345, -1.386753, -2.562567, -0.763069, 1.570796, 2.040141],accel_mss,speed_ms,0,blend_radius_m)
  movel([0.465719, -1.382944, -2.565284, -0.764161, 1.570796, 2.036515],accel_mss,speed_ms,0,blend_radius_m)
  movel([0.463468, -1.379991, -2.567376, -0.765022, 1.570796, 2.034264],accel_mss,speed_ms,0,blend_radius_m)
  movel([0.461113, -1.376292, -2.569979, -0.766117, 1.570796, 2.031910],accel_mss,speed_ms,0,blend_radius_m)
  movel([0.458810, -1.371807, -2.573109, -0.767472, 1.570796, 2.029607],accel_mss,speed_ms,0,blend_radius_m)
  movel([0.456708, -1.366486, -2.576786, -0.769117, 1.570796, 2.027504],accel_mss,speed_ms,0,blend_radius_m)
  movel([0.455614, -1.362516, -2.579504, -0.770370, 1.570796, 2.026411],accel_mss,speed_ms,0,blend_radius_m)
  movel([0.455031, -1.358689, -2.582102, -0.771598, 1.570796, 2.025827],accel_mss,speed_ms,0,blend_radius_m)
  movel([0.454907, -1.355018, -2.584575, -0.772796, 1.570796, 2.025703],accel_mss,speed_ms,0,blend_radius_m)
  movel([0.455182, -1.351514, -2.586918, -0.773957, 1.570796, 2.025978],accel_mss,speed_ms,0,blend_radius_m)
  movel([0.455800, -1.348197, -2.589121, -0.775071, 1.570796, 2.026596],accel_mss,speed_ms,0,blend_radius_m)
  movel([0.456698, -1.345080, -2.591177, -0.776132, 1.570796, 2.027495],accel_mss,speed_ms,0,blend_radius_m)
  movel([0.457819, -1.342179, -2.593078, -0.777132, 1.570796, 2.028615],accel_mss,speed_ms,0,blend_radius_m)
  movel([0.459097, -1.339513, -2.594815, -0.778060, 1.570796, 2.029894],accel_mss,speed_ms,0,blend_radius_m)
  movel([0.461874, -1.334952, -2.597765, -0.779672, 1.570796, 2.032671],accel_mss,speed_ms,0,blend_radius_m)
  movel([0.464513, -1.331530, -2.599960, -0.780899, 1.570796, 2.035309],accel_mss,speed_ms,0,blend_radius_m)
  movel([0.466479, -1.329387, -2.601326, -0.781676, 1.570796, 2.037275],accel_mss,speed_ms,0,blend_radius_m)
